// TwinCAT 3 PLC project otel
// Title: TcOtlp
// Company: S&E Engineering
// ProjectVersion: 0.0.0.1
// ProgramVersion: 3.1.4026.27
// libraries:
//   Tc2_Standard, * (Beckhoff Automation GmbH)
//   Tc2_System, * (Beckhoff Automation GmbH)
//   Tc2_Utilities, * (Beckhoff Automation GmbH)
//   Tc3_IotBase, * (Beckhoff Automation GmbH)
//   Tc3_JsonXml, * (Beckhoff Automation GmbH)
// project tree:
//   OTEL/COMMON/ENUMS/ E_BytesEncoding.TcTLEO
//   OTEL/COMMON/FUNCTION_BLOCKS/ FB_InstrumentationScope.TcPOU, FB_Resource.TcPOU
//   OTEL/COMMON/STRUCTS/ ST_LinkedListNode.TcDUT
//   OTEL/EXPORTING/ENUMS/ E_FileExporterState.TcTLEO, E_HttpExporterState.TcTLEO
//   OTEL/LOGGING/EXPORTING/ENUMS/ E_LogRecordExporterFailureReason.TcTLEO, E_LogRecordExporterState.TcTLEO
//   OTEL/LOGGING/EXPORTING/FUNCTION_BLOCKS/ FB_LogRecordExporter_Base.TcPOU, FB_LogRecordExporter_Console.TcPOU, FB_LogRecordExporter_File.TcPOU, FB_LogRecordExporter_HTTP.TcPOU
//   OTEL/LOGGING/LOGGER/ENUMS/ E_LoggerFailureReason.TcTLEO
//   OTEL/LOGGING/LOGGER/FUNCTION_BLOCKS/ FB_Logger.TcPOU
//   OTEL/LOGGING/LOG_RECORD/ENUMS/ E_LogRecordCloneFailureReason.TcTLEO, E_LogRecordFlag.TcTLEO, E_LogRecordQueueFailureReason.TcTLEO, E_SeverityNumber.TcTLEO
//   OTEL/LOGGING/LOG_RECORD/FUNCTION_BLOCKS/ FB_LogRecord.TcPOU, FB_LogRecordQueue.TcPOU
//   OTEL/LOGGING/PROCESSORS/ENUMS/ E_LogRecordProcessorFailureReason.TcTLEO
//   OTEL/LOGGING/PROCESSORS/FUNCTION_BLOCKS/ FB_LogRecordProcessor_Base.TcPOU, FB_LogRecordProcessor_Batch.TcPOU, FB_LogRecordProcessor_Simple.TcPOU
//   OTEL/LOGGING/PROVIDER/ENUMS/ E_LoggerProviderFailureReason.TcTLEO
//   OTEL/LOGGING/PROVIDER/FUNCTION_BLOCKS/ FB_LoggerProvider.TcPOU
//   OTEL/LOGGING/SERIALIZATION/FUNCTION_BLOCKS/ FB_LogRecordProtoJsonSerializer.TcPOU
//   OTEL/ TcOtlp_GVL.TcGVL
//   OTEL/TRACING/EXPORTING/ENUMS/ E_SpanExporterFailureReason.TcTLEO
//   OTEL/TRACING/EXPORTING/FUNCTION_BLOCKS/ FB_SpanExporter_Base.TcPOU, FB_SpanExporter_File.TcPOU, FB_SpanExporter_Console.TcPOU, FB_SpanExporter_HTTP.TcPOU
//   OTEL/TRACING/SPAN/ENUMS/ E_SpanCloneFailureReason.TcTLEO, E_SpanFlags.TcTLEO, E_ContextFactoryFailureReason.TcTLEO, E_SpanKind.TcTLEO, E_SpanQueueFailureReason.TcTLEO, E_StatusCode.TcTLEO
//   OTEL/TRACING/PROCESSORS/ENUMS/ E_SpanProcessorFailureReason.TcTLEO
//   OTEL/TRACING/PROCESSORS/FUNCTION_BLOCKS/ FB_SpanProcessor_Batch.TcPOU, FB_SpanProcessor_Base.TcPOU, FB_SpanProcessor_Simple.TcPOU
//   OTEL/EXPORTING/STRUCTS/ ST_HttpEndpoint.TcDUT
//   OTEL/EXPORTING/FUNCTIONS/ F_ParseHttpUrl.TcPOU
//   OTEL/TRACING/TRACESTATE/ENUMS/ E_TraceStateFailureReason.TcTLEO
//   OTEL/TRACING/TRACESTATE/FUNCTION_BLOCKS/ FB_TraceState.TcPOU, TraceStateFactory.TcPOU
//   OTEL/TRACING/PROPAGATION/ENUMS/ E_PropagationFailureReason.TcTLEO
//   OTEL/TRACING/PROPAGATION/ TraceContextPropagator.TcPOU
//   OTEL/TRACING/PROPAGATION/STRUCTS/ ST_TraceContextCarrier.TcDUT
//   OTEL/TRACING/SAMPLING/FUNCTION_BLOCKS/ FB_Sampler.TcPOU, FB_Sampler_AlwaysOn.TcPOU, FB_Sampler_ErrorsOnly.TcPOU
//   OTEL/TRACING/ID_GENERATION/ENUMS/ E_IdGenFailureReason.TcTLEO
//   OTEL/TRACING/ID_GENERATION/FUNCTION_BLOCKS/ FB_IdGenerator.TcPOU, FB_IdGenerator_Base.TcPOU
//   OTEL/TRACING/LINK/ENUM/ E_LinkFailureReason.TcTLEO
//   OTEL/TRACING/LINK/FUNCTION_BLOCKS/ FB_Link.TcPOU, FB_Links.TcPOU, LinkFactory.TcPOU
//   OTEL/TRACING/PROVIDER/ENUMS/ E_TracerProviderFailureReason.TcTLEO
//   OTEL/TRACING/PROVIDER/FUNCTION_BLOCKS/ FB_TracerProvider.TcPOU
//   OTEL/TRACING/SERIALIZATION/FUNCTION_BLOCKS/ FB_SpanProtoJsonSerializer.TcPOU
//   OTEL/TRACING/SPAN/ ContextFactory.TcPOU
//   OTEL/TRACING/SPAN/FUNCTION_BLOCKS/ FB_Span.TcPOU, FB_SpanContext.TcPOU, FB_SpanQueue.TcPOU, FB_Status.TcPOU
//   OTEL/TRACING/TRACER/ENUMS/ E_TracerFailureReason.TcTLEO
//   OTEL/TRACING/TRACER/ FB_Tracer.TcPOU
//   OTEL/VALUES/ENUMS/ E_AttributesFailureReason.TcTLEO, E_ValueFactoryFailureReason.TcTLEO, E_ValueType.TcTLEO
//   OTEL/VALUES/FUNCTION_BLOCKS/ FB_AnyValue.TcPOU, FB_Attributes.TcPOU, FB_KeyValue.TcPOU, FB_Number.TcPOU, FB_SpanId.TcPOU, FB_String.TcPOU, FB_TraceId.TcPOU
//   OTEL/VALUES/INTERFACES/ I_OtlpValue.TcIO
//   OTEL/VALUES/ ValueFactory.TcPOU
//   OTEL/SERIALIZATION/FUNCTION_BLOCKS/ FB_BaseProtoJsonSerializer.TcPOU
//   OTEL/SERIALIZATION/ENUMS/ E_ProtoJsonSerializerFailureReason.TcTLEO
//   Project Information/ F_GetCompany.TcPOU, F_GetTitle.TcPOU, F_GetVersion.TcPOU
//   Version/ Global_Version.TcGVL
// (motion and I/O tree: see PLC project test)
// real-time tasks:
//   TASK PlcTask: cycle T#10ms, priority 20, ADS port 350

// ---- OTEL/COMMON/ENUMS/E_BytesEncoding.TcTLEO
{attribute 'qualified_only'}
{attribute 'strict'}
{attribute 'to_string'}
TYPE E_BytesEncoding :
(
	hex := 0,
	base64
);
END_TYPE

// ---- OTEL/COMMON/STRUCTS/ST_LinkedListNode.TcDUT
{attribute 'enable_dynamic_creation'}
TYPE ST_LinkedListNode :
STRUCT
	val: PVOID;
	nxt: POINTER TO ST_LinkedListNode;
END_STRUCT
END_TYPE

// ---- OTEL/EXPORTING/ENUMS/E_FileExporterState.TcTLEO
{attribute 'qualified_only'}
{attribute 'strict'}
{attribute 'to_string'}
TYPE E_FileExporterState :
(
	error := -10,
	idle := 0,
	serializing := 10,
	creating := 15,
	opening := 20,
	buffering := 25,
	writing := 30,
	closing := 40,
	rotating := 50,
	done := 99
);
END_TYPE
//  error = '-10'

// ---- OTEL/EXPORTING/ENUMS/E_HttpExporterState.TcTLEO
{attribute 'qualified_only'}
{attribute 'strict'}
{attribute 'to_string'}
TYPE E_HttpExporterState :
(
	error := -10,
	idle := 0,
	serializing := 10,
	sending := 20,
	waiting := 30,
	processing := 40,
	done := 99
);
END_TYPE
//  error = '-10'

// ---- OTEL/LOGGING/EXPORTING/ENUMS/E_LogRecordExporterFailureReason.TcTLEO
{attribute 'qualified_only'}
{attribute 'strict'}
{attribute 'to_string'}
TYPE E_LogRecordExporterFailureReason :
(
	NA := 0,  // No failure occurred.
	ACTIVE_EXPORT_IN_PROGRESS,  // The exporter cannot accept another batch while an export is active.
	QUEUE_TRANSFER_FAILURE,  // Records could not be transferred into the exporter queue.
	SERIALIZATION_FAILURE,  // The accepted records could not be serialized.
	BUFFER_ALLOCATION_FAILURE,  // The serialized payload buffer could not be allocated.
	FILE_OPEN_FAILURE,  // The destination file could not be opened.
	FILE_WRITE_FAILURE,  // The serialized payload could not be written.
	FILE_CLOSE_FAILURE,  // The destination file could not be closed.
	HTTP_URL_PARSE_FAILURE,  // The configured endpoint URL could not be parsed.
	HTTP_REQUEST_FAILURE,  // The HTTP request could not be sent or completed.
	HTTP_STATUS_FAILURE  // The server responded with a non-success HTTP status code.
) UDINT;
END_TYPE

// ---- OTEL/LOGGING/EXPORTING/ENUMS/E_LogRecordExporterState.TcTLEO
{attribute 'qualified_only'}
{attribute 'strict'}
{attribute 'to_string'}
TYPE E_LogRecordExporterState :
(
	SUCCESS := 0,
	BUSY,
	FAILURE
);
END_TYPE

// ---- OTEL/LOGGING/LOGGER/ENUMS/E_LoggerFailureReason.TcTLEO
{attribute 'qualified_only'}
{attribute 'strict'}
{attribute 'to_string'}
TYPE E_LoggerFailureReason :
(
	NA := 0,  // No failure occurred.
	LOG_RECORD_ALREADY_STARTED,  // A record is already being built by this logger.
	LOG_RECORD_NOT_STARTED,  // No active record is available to modify or emit.
	EVENT_NAME_INVALID,  // The event name could not be copied into an owned value.
	BODY_VALUE_POINTER_NULL,  // The supplied body value pointer is null.
	BODY_VALUE_INVALID,  // The supplied body value could not be cloned.
	BODY_VALUE_TYPE_UNSUPPORTED,  // The supplied body value type is not supported.
	ATTRIBUTE_VALUE_INVALID,  // An attribute could not be created from the supplied value.
	ATTRIBUTE_VALUE_TYPE_UNSUPPORTED,  // The supplied attribute value type is not supported.
	ATTRIBUTE_COUNT_LIMIT_REACHED,  // The record cannot own another attribute.
	SPAN_ID_BYTES_POINTER_NULL,  // The supplied Span ID byte pointer is null.
	SPAN_ID_BYTE_COUNT_TOO_SMALL,  // The supplied Span ID buffer is shorter than eight bytes.
	SPAN_ID_INVALID,  // The supplied Span ID could not be copied.
	TRACE_ID_BYTES_POINTER_NULL,  // The supplied Trace ID byte pointer is null.
	TRACE_ID_BYTE_COUNT_TOO_SMALL,  // The supplied Trace ID buffer is shorter than sixteen bytes.
	TRACE_ID_INVALID,  // The supplied Trace ID could not be copied.
	SNAPSHOT_COPY_FAILURE,  // The resource or instrumentation-scope snapshot could not be copied.
	MEMORY_ALLOCATION_FAILURE,  // Dynamic memory allocation failed.
	TRANSFER_TO_PROVIDER_FAILURE  // Could not transfer ownership of the record to the provider
) UDINT;
END_TYPE

// ---- OTEL/LOGGING/LOG_RECORD/ENUMS/E_LogRecordCloneFailureReason.TcTLEO
{attribute 'qualified_only'}
{attribute 'strict'}
{attribute 'to_string'}
TYPE E_LogRecordCloneFailureReason :
(
	NA := 0,  // No failure occurred.
	DESTINATION_ALREADY_ASSIGNED,  // The clone destination pointer is already assigned.
	EVENT_NAME_INVALID,  // The source event name could not be cloned.
	TRACE_ID_INVALID,  // The source Trace ID could not be cloned.
	SPAN_ID_INVALID,  // The source Span ID could not be cloned.
	BODY_VALUE_INVALID,  // The source body could not be cloned.
	BODY_VALUE_TYPE_UNSUPPORTED,  // The source body contains an unsupported value type.
	RESOURCE_COPY_FAILURE,  // The resource snapshot could not be copied.
	SCOPE_COPY_FAILURE,  // The instrumentation-scope snapshot could not be copied.
	ATTRIBUTE_COPY_FAILURE,  // The record attributes could not be copied.
	MEMORY_ALLOCATION_FAILURE  // Dynamic memory allocation failed.
) UDINT;
END_TYPE

// ---- OTEL/LOGGING/LOG_RECORD/ENUMS/E_LogRecordFlag.TcTLEO
{attribute 'qualified_only'}
{attribute 'strict'}
{attribute 'to_string'}
TYPE E_LogRecordFlag:
(
	// The zero value for the enum. Should not be used for comparisons.
	// Instead use bitwise "and" with the appropriate mask as shown above.
	LOG_RECORD_FLAGS_DO_NOT_USE := 0,
	// Bits 0-7 are used for trace flags.
	LOG_RECORD_FLAGS_TRACE_FLAGS_MASK := 255 //0x000000FF;
) UDINT;
END_TYPE
//  LOG_RECORD_FLAGS_TRACE_FLAGS_MASK = '255 '

// ---- OTEL/LOGGING/LOG_RECORD/ENUMS/E_LogRecordQueueFailureReason.TcTLEO
{attribute 'qualified_only'}
{attribute 'strict'}
{attribute 'to_string'}
TYPE E_LogRecordQueueFailureReason :
(
	NA := 0,  // No failure occurred.
	RECORD_POINTER_NULL,  // The supplied log-record pointer is null.
	DESTINATION_ALREADY_ASSIGNED,  // The pop destination pointer is already assigned.
	QUEUE_EMPTY,  // The queue contains no record to pop.
	MAX_SIZE_ENFORCEMENT_FAILURE := 5,  // The bounded eviction loop could not restore the configured maximum size.
	DESTINATION_NOT_EMPTY,  // The transfer destination already owns records.
	DESTINATION_CAPACITY_TOO_SMALL,  // The transfer destination cannot hold every source record.
	SELF_TRANSFER_NOT_ALLOWED,  // A queue cannot transfer ownership to itself.
	MEMORY_ALLOCATION_FAILURE  // Dynamic node allocation failed.
) UDINT;
END_TYPE

// ---- OTEL/LOGGING/LOG_RECORD/ENUMS/E_SeverityNumber.TcTLEO
{attribute 'qualified_only'}
{attribute 'strict'}
{attribute 'to_string'}
TYPE E_SeverityNumber :
(
	UNSPECIFIED := 0,
	TRACE,
	TRACE2,
	TRACE3,
	TRACE4,
	DEBUG,
	DEBUG2,
	DEBUG3,
	DEBUG4,
	INFO,
	INFO2,
	INFO3,
	INFO4,
	WARN,
	WARN2,
	WARN3,
	WARN4,
	ERROR,
	ERROR2,
	ERROR3,
	ERROR4,
	FATAL,
	FATAL2,
	FATAL3,
	FATAL4
);
END_TYPE

// ---- OTEL/LOGGING/PROCESSORS/ENUMS/E_LogRecordProcessorFailureReason.TcTLEO
{attribute 'qualified_only'}
{attribute 'strict'}
{attribute 'to_string'}
TYPE E_LogRecordProcessorFailureReason :
(
	NA := 0,  // No failure occurred.
	RECORD_CLONE_FAILURE,  // The emitted record could not be cloned for retention.
	QUEUE_PUSH_FAILURE,  // The retained record could not be transferred into the queue.
	EXPORT_FAILURE  // The exporter did not accept the prepared batch.
) UDINT;
END_TYPE

// ---- OTEL/LOGGING/PROVIDER/ENUMS/E_LoggerProviderFailureReason.TcTLEO
{attribute 'qualified_only'}
{attribute 'strict'}
{attribute 'to_string'}
TYPE E_LoggerProviderFailureReason :
(
	NA := 0,  // No failure occurred.
	RECORD_POINTER_NULL,  // The supplied log record pointer is null.
	QUEUE_POP_FAILURE,  // A record could not be popped from the provider's queue during cyclical processing.
	STAGE_PROCESSOR_FAILURE,  // A processor could not be added to the internal linked list for some reason.
	UNEXPECTED_NULL_PROCESSOR_POINTER,  // A processor pointer was invalid when being accessed internally to the provider.
	UNEXPECTED_NULL_LINKED_LIST_NODE  // A processor linked list poitner was invalid when being accessed internally to the provider.
) UDINT;
END_TYPE

// ---- OTEL/TRACING/EXPORTING/ENUMS/E_SpanExporterFailureReason.TcTLEO
(* Why a span exporter refused a batch or could not deliver it. *)
{attribute 'qualified_only'}
{attribute 'strict'}
{attribute 'to_string'}
TYPE E_SpanExporterFailureReason :
(
	NA := 0,  // No failure occurred.
	ACTIVE_EXPORT_IN_PROGRESS,  // The exporter cannot accept another batch while an export is active.
	QUEUE_TRANSFER_FAILURE,  // Spans could not be transferred into the exporter queue.
	SERIALIZATION_FAILURE,  // The accepted spans could not be serialized.
	BUFFER_ALLOCATION_FAILURE,  // The serialized payload buffer could not be allocated.
	FILE_OPEN_FAILURE,  // The destination file could not be opened.
	FILE_WRITE_FAILURE,  // The serialized payload could not be written.
	FILE_CLOSE_FAILURE,  // The destination file could not be closed.
	HTTP_URL_PARSE_FAILURE,  // The configured endpoint URL could not be parsed.
	HTTP_REQUEST_FAILURE,  // The HTTP request could not be sent or completed.
	HTTP_STATUS_FAILURE  // The server responded with a non-success HTTP status code.
) UDINT;
END_TYPE

// ---- OTEL/TRACING/SPAN/ENUMS/E_SpanCloneFailureReason.TcTLEO
(* Why FB_Span.cloneTo could not copy a span. *)
{attribute 'qualified_only'}
{attribute 'strict'}
{attribute 'to_string'}
TYPE E_SpanCloneFailureReason :
(
	NA := 0,  // No failure occurred.
	DESTINATION_ALREADY_ASSIGNED,  // The destination pointer was not 0.
	MEMORY_ALLOCATION_FAILURE,  // Dynamic memory allocation failed.
	VALUE_COPY_FAILURE,  // The name, an identifier, the trace state or the status message could not be copied.
	ATTRIBUTE_COPY_FAILURE,  // The span attributes could not be copied.
	LINK_COPY_FAILURE,  // A span link could not be copied.
	RESOURCE_COPY_FAILURE,  // The resource could not be copied.
	SCOPE_COPY_FAILURE  // The instrumentation scope could not be copied.
) UDINT;
END_TYPE

// ---- OTEL/TRACING/PROCESSORS/ENUMS/E_SpanProcessorFailureReason.TcTLEO
(* Why a span processor could not keep or export an ended span. *)
{attribute 'qualified_only'}
{attribute 'strict'}
{attribute 'to_string'}
TYPE E_SpanProcessorFailureReason :
(
	NA := 0,  // No failure occurred.
	SPAN_CLONE_FAILURE,  // The ended span could not be cloned for retention.
	QUEUE_PUSH_FAILURE,  // The clone could not be pushed onto the queue.
	EXPORT_FAILURE  // The exporter did not accept the prepared batch.
) UDINT;
END_TYPE

// ---- OTEL/EXPORTING/STRUCTS/ST_HttpEndpoint.TcDUT
(* An HTTP endpoint split out of a URL by F_ParseHttpUrl. *)
TYPE ST_HttpEndpoint :
STRUCT
	useTls: BOOL;  // TRUE for https
	host: T_MaxString;
	port: UINT;  // the explicit port, or 80 for http and 443 for https
	path: T_MaxString := '/';  // starts with '/'
END_STRUCT
END_TYPE

// ---- OTEL/TRACING/TRACESTATE/ENUMS/E_TraceStateFailureReason.TcTLEO
(* Why TraceStateFactory could not produce a trace state. *)
{attribute 'qualified_only'}
{attribute 'strict'}
{attribute 'to_string'}
TYPE E_TraceStateFailureReason :
(
	NA := 0,  // No failure.
	DESTINATION_ALREADY_ASSIGNED,  // The destination pointer already holds a trace state.
	SOURCE_POINTER_NULL,  // The source trace state is missing or has been freed.
	HEADER_POINTER_NULL,  // The header pointer is 0.
	HEADER_TOO_LONG,  // The header is longer than TraceStateFactory.MAX_HEADER_LENGTH.
	INVALID_KEY,  // An entry has a key that does not follow the W3C key grammar.
	INVALID_VALUE,  // An entry has no '=' or a value that does not follow the W3C value grammar.
	DUPLICATE_KEY,  // Two entries have the same key.
	TOO_MANY_ENTRIES,  // The header has more than TraceStateFactory.MAX_ENTRIES entries.
	MEMORY_ALLOCATION_FAILURE  // The trace state could not be allocated.
) UDINT;
END_TYPE

// ---- OTEL/TRACING/PROPAGATION/ENUMS/E_PropagationFailureReason.TcTLEO
(* Why TraceContextPropagator could not extract a span context from a carrier, or inject one into it. *)
{attribute 'qualified_only'}
{attribute 'strict'}
{attribute 'to_string'}
TYPE E_PropagationFailureReason :
(
	NA := 0,  // No failure.
	DESTINATION_ALREADY_ASSIGNED,  // The destination pointer already holds a span context.
	TRACEPARENT_EMPTY,  // No traceparent arrived, so there is no context to extract.
	TRACEPARENT_LENGTH_INVALID,  // The traceparent is shorter than 55 characters, or longer for version 00.
	VERSION_INVALID,  // The version is not two lowercase hex digits, or is the reserved ff.
	DELIMITER_INVALID,  // A field is not followed by '-', or a future version's flags are followed by something else.
	TRACE_ID_INVALID,  // The trace id is not 32 lowercase hex digits, or is all zero.
	SPAN_ID_INVALID,  // The parent span id is not 16 lowercase hex digits, or is all zero.
	TRACE_FLAGS_INVALID,  // The trace flags are not two lowercase hex digits.
	MEMORY_ALLOCATION_FAILURE,  // The span context, or a shortened trace state, could not be allocated.
	CONTEXT_POINTER_NULL,  // inject was given no span context.
	CONTEXT_INVALID  // The span context has an all-zero trace id or span id, so there is nothing to propagate.
) UDINT;
END_TYPE

// ---- OTEL/TRACING/PROPAGATION/STRUCTS/ST_TraceContextCarrier.TcDUT
(*
	The W3C Trace Context headers of one call, written by TraceContextPropagator.inject and read
	by extract. It is the contract between the propagator and a transport: a transport moves the
	whole block, so the receiver never sees a traceparent beside a stale tracestate, and it knows
	nothing about the headers' format. The traceparent fits version 00, and the tracestate fits
	the 512 characters W3C asks every vendor to propagate.
*)
TYPE ST_TraceContextCarrier :
STRUCT
	traceparent: STRING(55);
	tracestate: STRING(512);  // '' when the context has no trace state
END_STRUCT
END_TYPE

// ---- OTEL/TRACING/ID_GENERATION/ENUMS/E_IdGenFailureReason.TcTLEO
{attribute 'qualified_only'}
{attribute 'strict'}
{attribute 'to_string'}
TYPE E_IdGenFailureReason :
(
	NA := 0,  // No failure occurred.
	NO_IDENTIFIERS_AVAILABLE,  // The ring held too few bytes; the caller must retry on a later cycle.
	GUID_SERVICE_FAILED,  // The TwinCAT GUID service reported an error while the ring was being refilled.
	MEMORY_ALLOCATION_FAILURE,  // The ring could not be allocated.
	INVALID_CONFIGUATION  // parameters used to configure the generator were not valid
) UDINT;
END_TYPE

// ---- OTEL/TRACING/LINK/ENUM/E_LinkFailureReason.TcTLEO
(* Why a LinkFactory or FB_Links call failed. *)
{attribute 'qualified_only'}
{attribute 'strict'}
{attribute 'to_string'}
TYPE E_LinkFailureReason :
(
	NA := 0,  // No failure occurred.
	DESTINATION_ALREADY_ASSIGNED,  // The destination pointer was not 0.
	CONTEXT_POINTER_NULL,  // The span context pointer is null.
	CONTEXT_INVALID,  // The span context has an all zero trace id or span id.
	SPAN_POINTER_NULL,  // The span pointer is null.
	LINK_POINTER_NULL,  // The link pointer is null.
	LINK_COUNT_LIMIT_REACHED,  // The collection already holds maxCount links; the link was dropped and counted.
	LINKS_EMPTY,  // The collection holds no links.
	MEMORY_ALLOCATION_FAILURE,  // Dynamic memory allocation failed.
	ATTRIBUTE_COPY_FAILURE  // The link attributes could not be copied.
) UDINT;
END_TYPE

// ---- OTEL/TRACING/PROVIDER/ENUMS/E_TracerProviderFailureReason.TcTLEO
(* Why FB_TracerProvider.tick failed. *)
{attribute 'qualified_only'}
{attribute 'strict'}
{attribute 'to_string'}
TYPE E_TracerProviderFailureReason :
(
	NA := 0,  // No failure occurred.
	QUEUE_POP_FAILURE,  // An ended span could not be popped from the provider queue.
	STAGE_PROCESSOR_FAILURE,  // A processor could not be added to the staged list.
	UNEXPECTED_NULL_PROCESSOR_POINTER,  // A staged processor pointer was null.
	UNEXPECTED_NULL_LINKED_LIST_NODE,  // The staged list was shorter than stagedProcessorCount.
	ID_GENERATOR_TICK_FAILURE  // The id generator could not advance.
) UDINT;
END_TYPE

// ---- OTEL/TRACING/SPAN/ENUMS/E_SpanFlags.TcTLEO
{attribute 'qualified_only'}
{attribute 'strict'}
{attribute 'to_string'}
TYPE E_SpanFlags :
(
	// The zero value for the enum. Should not be used for comparisons.
	// Instead use bitwise "and" with the appropriate mask as shown above.
	SPAN_FLAGS_DO_NOT_USE := 16#0,

	// Bits 0-7 are used for trace flags.
	SPAN_FLAGS_TRACE_FLAGS_MASK := 16#000000FF,

	// Bits 8 and 9 are used to indicate that the parent span or link span is remote.
	// Bit 8 (`HAS_IS_REMOTE`) indicates whether the value is known.
	// Bit 9 (`IS_REMOTE`) indicates whether the span or link is remote.
	SPAN_FLAGS_CONTEXT_HAS_IS_REMOTE_MASK := 16#00000100,
	SPAN_FLAGS_CONTEXT_IS_REMOTE_MASK := 16#00000200

  // Bits 10-31 are reserved for future use.
) UDINT;
END_TYPE
//  SPAN_FLAGS_DO_NOT_USE = '16#0'
//  SPAN_FLAGS_TRACE_FLAGS_MASK = '16#000000FF'
//  SPAN_FLAGS_CONTEXT_HAS_IS_REMOTE_MASK = '16#00000100'
//  SPAN_FLAGS_CONTEXT_IS_REMOTE_MASK = '16#00000200  '

// ---- OTEL/TRACING/SPAN/ENUMS/E_ContextFactoryFailureReason.TcTLEO
{attribute 'qualified_only'}
{attribute 'strict'}
{attribute 'to_string'}
TYPE E_ContextFactoryFailureReason :
(
	NA := 0,  // No failure occurred.
	DESTINATION_ALREADY_ASSIGNED,  // The destination pointer was already assigned when the operation began.
	TRACE_ID_POINTER_NULL,  // The trace ID pointer is null.
	SPAN_ID_POINTER_NULL,  // The span ID pointer is null.
	MEMORY_ALLOCATION_FAILURE,  // Dynamic memory allocation failed.
	SPAN_POINTER_NULL  // fromSpan was given a null span pointer.
);
END_TYPE

// ---- OTEL/TRACING/SPAN/ENUMS/E_SpanKind.TcTLEO
{attribute 'qualified_only'}
{attribute 'strict'}
{attribute 'to_string'}
TYPE E_SpanKind :
(
	// Unspecified. Do NOT use as default.
	// Implementations MAY assume SpanKind to be INTERNAL when receiving UNSPECIFIED.
	SPAN_KIND_UNSPECIFIED := 0,
	
	// Indicates that the span represents an internal operation within an application,
	// as opposed to an operation happening at the boundaries. Default value.
	SPAN_KIND_INTERNAL := 1,
	
	// Indicates that the span covers server-side handling of an RPC or other
	// remote network request.
	SPAN_KIND_SERVER := 2,
	
	// Indicates that the span describes a request to some remote service.
	SPAN_KIND_CLIENT := 3,
	
	// Indicates that the span describes a producer sending a message to a broker.
	// Unlike CLIENT and SERVER, there is often no direct critical path latency relationship
	// between producer and consumer spans. A PRODUCER span ends when the message was accepted
	// by the broker while the logical processing of the message might span a much longer time.
	SPAN_KIND_PRODUCER := 4,
	
	// Indicates that the span describes consumer receiving a message from a broker.
	// Like the PRODUCER kind, there is often no direct critical path latency relationship
	// between producer and consumer spans.
	SPAN_KIND_CONSUMER := 5
) UDINT;
END_TYPE

// ---- OTEL/TRACING/SPAN/ENUMS/E_SpanQueueFailureReason.TcTLEO
{attribute 'qualified_only'}
{attribute 'strict'}
{attribute 'to_string'}
TYPE E_SpanQueueFailureReason :
(
	NA := 0,  // No failure occurred.
	SPAN_POINTER_NULL,  // The supplied span pointer is null.
	DESTINATION_ALREADY_ASSIGNED,  // The pop destination pointer is already assigned.
	QUEUE_EMPTY,  // The queue contains no span to pop.
	MAX_SIZE_ENFORCEMENT_FAILURE,  // The bounded eviction loop could not restore the configured maximum size.
	MEMORY_ALLOCATION_FAILURE,  // Dynamic node allocation failed.
	SELF_TRANSFER_NOT_ALLOWED,  // transferTo was asked to move spans into the same queue.
	DESTINATION_NOT_EMPTY  // transferTo needs an empty destination queue.
) UDINT;
END_TYPE

// ---- OTEL/TRACING/SPAN/ENUMS/E_StatusCode.TcTLEO
{attribute 'qualified_only'}
{attribute 'strict'}
{attribute 'to_string'}
TYPE E_StatusCode :
(
	// The default status.
	STATUS_CODE_UNSET := 0,
	// The Span has been validated by an Application developer or Operator to 
	// have completed successfully.
	STATUS_CODE_OK := 1,
	// The Span contains an error.
	STATUS_CODE_ERROR := 2
) UDINT;
END_TYPE

// ---- OTEL/TRACING/TRACER/ENUMS/E_TracerFailureReason.TcTLEO
{attribute 'qualified_only'}
{attribute 'strict'}
{attribute 'to_string'}
TYPE E_TracerFailureReason :
(
	NA := 0,  // No failure occurred.
	SPAN_ALREADY_STARTED,  // startSpan was called while a span was still being built.
	SPAN_NOT_STARTED,  // No span is being built to modify or hand over.
	SPAN_NAME_EMPTY,  // The span name is empty.
	SPAN_KIND_UNSPECIFIED,  // SPAN_KIND_UNSPECIFIED was given; OTLP says not to use it.
	PARENT_CONTEXT_POINTER_NULL,  // The parent context pointer is null.
	PARENT_CONTEXT_INVALID,  // The parent context has an all zero trace id or span id.
	ATTRIBUTE_VALUE_INVALID,  // An attribute could not be created from the supplied value.
	ATTRIBUTE_VALUE_TYPE_UNSUPPORTED,  // The supplied attribute value type is not supported.
	ATTRIBUTE_COUNT_LIMIT_REACHED,  // The span cannot own another attribute.
	DESTINATION_ALREADY_ASSIGNED,  // The destination pointer was already assigned when build began.
	IDENTIFIERS_UNAVAILABLE,  // The id generator had no identifiers ready; retry on a later cycle.
	ID_GENERATION_FAILURE,  // The id generator failed for another reason.
	SNAPSHOT_COPY_FAILURE,  // The resource or instrumentation-scope snapshot could not be copied.
	MEMORY_ALLOCATION_FAILURE,  // Dynamic memory allocation failed.
	SPAN_POINTER_NULL,  // A method for a running span, such as endSpan, was given a null span pointer.
	TRANSFER_TO_PROVIDER_FAILURE,  // The provider could not queue the ended span, so it was released.
	LINK_CONTEXT_POINTER_NULL,  // addLink was given a null span context pointer.
	LINK_CONTEXT_INVALID,  // The linked context has an all zero trace id or span id.
	LINK_COUNT_LIMIT_REACHED,  // The span cannot own another link.
	PARENT_SPAN_POINTER_NULL,  // setParentUsingSpan was given a null span pointer.
	PARENT_SPAN_INVALID,  // The parent span has not been built, so it has no trace id or span id.
	SPAN_STATUS_ALREADY_SET,  // The span already has a status, and the first one set wins.
	SPAN_INVALID,  // The span has not been built, so it has no trace id or span id.
	LINK_POINTER_NULL  // pushSpanLink was given a null link pointer.
) UDINT;
END_TYPE

// ---- OTEL/VALUES/ENUMS/E_AttributesFailureReason.TcTLEO
{attribute 'qualified_only'}
{attribute 'strict'}
{attribute 'to_string'}
TYPE E_AttributesFailureReason :
(
	NA := 0,  // No attribute failure occurred.
	KV_POINTER_NULL,  // The supplied key-value pair pointer is null.
	KV_KEY_POINTER_NULL,  // The key-value pair has no key.
	KV_VALUE_POINTER_NULL,  // The key-value pair has no value.
	KV_VALUE_INVALID,  // The key-value pair contains an invalid value.
	KV_VALUE_TYPE_UNSUPPORTED,  // The key-value pair contains an unsupported value type.
	ATTRIBUTE_COUNT_LIMIT_REACHED,  // Adding a new key would exceed the configured attribute count limit.
	MEMORY_ALLOCATION_FAILURE,  // Dynamic memory allocation failed.
	KEY_NOT_FOUND  // The source collection has no attribute with the requested key.
) UDINT;
END_TYPE

// ---- OTEL/VALUES/ENUMS/E_ValueFactoryFailureReason.TcTLEO
{attribute 'qualified_only'}
{attribute 'strict'}
{attribute 'to_string'}
TYPE E_ValueFactoryFailureReason :
(
	NA := 0,  // No failure occurred.
	DESTINATION_ALREADY_ASSIGNED,  // The destination pointer was already assigned when the operation began.
	SOURCE_POINTER_NULL,  // The source pointer is null.
	NUMBER_VALUE_POINTER_NULL,  // The numeric value pointer is null.
	NUMBER_VALUE_SIZE_INVALID,  // The numeric value size is zero or negative.
	KEY_POINTER_NULL,  // The key pointer is null.
	VALUE_POINTER_NULL,  // The value pointer is null.
	STRING_POINTER_NULL,  // The string pointer is null.
	SPAN_ID_BYTES_POINTER_NULL,  // The Span ID byte-array pointer is null.
	SPAN_ID_BYTE_COUNT_TOO_SMALL,  // The supplied byte count is too small for a Span ID.
	TRACE_ID_BYTES_POINTER_NULL,  // The Trace ID byte-array pointer is null.
	TRACE_ID_BYTE_COUNT_TOO_SMALL,  // The supplied byte count is too small for a Trace ID.
	UNSUPPORTED_VALUE_TYPE,  // The source value type is not supported by the factory operation.
	MEMORY_ALLOCATION_FAILURE  // Dynamic memory allocation failed.
);
END_TYPE

// ---- OTEL/VALUES/ENUMS/E_ValueType.TcTLEO
{attribute 'qualified_only'}
{attribute 'strict'}
{attribute 'to_string'}
TYPE E_ValueType :
(
	E_String := 0,
	E_TraceId,
	E_SpanId,
	E_AnyValue,
	E_KeyValue,
	E_Number
);
END_TYPE

// ---- OTEL/SERIALIZATION/ENUMS/E_ProtoJsonSerializerFailureReason.TcTLEO
{attribute 'qualified_only'}
{attribute 'strict'}
{attribute 'to_string'}
TYPE E_ProtoJsonSerializerFailureReason :
(
	NA := 0,  // No failure occurred.
	JSON_VALUE_INVALID,  // The destination JSON value is invalid.
	JSON_OPERATION_FAILURE,  // The JSON DOM parser could not create or append a value.
	KEY_POINTER_NULL,  // The supplied member-key pointer is null.
	VALUE_POINTER_NULL,  // The supplied OTLP value pointer is null.
	LOG_RECORD_POINTER_NULL,  // The supplied log-record pointer is null.
	NUMBER_VALUE_POINTER_NULL,  // The numeric value does not point to its concrete value.
	UNSUPPORTED_VALUE_TYPE,  // The OTLP value type is not supported.
	UNSUPPORTED_NUMBER_TYPE,  // The IEC numeric type is not supported.
	BYTES_POINTER_NULL,  // The byte-array pointer is null.
	BYTE_COUNT_ZERO,  // No bytes were supplied for encoding.
	STRING_POINTER_NULL,  // The destination or source string pointer is null.
	STRING_BUFFER_TOO_SMALL,  // The encoded value does not fit in the destination string.
	UNSUPPORTED_BYTES_ENCODING,  // The requested byte encoding is not supported.
	ATTRIBUTE_COLLECTION_INCONSISTENT,  // The attribute count and linked values disagree.
	LOG_RECORD_COLLECTION_INCONSISTENT,  // The queue count and linked records disagree.
	QUEUE_TRANSFER_FAILURE,  // Ownership could not be transferred to the serializer queue.
	QUEUE_POP_FAILURE,  // An owned record could not be removed from the serializer queue.
	QUEUE_ROTATE_FAILURE,  // The serializer queue could not preserve grouping order.
	LOOP_LIMIT_EXCEEDED,  // Serialization could not complete within GVL.MAX_LOOP_COUNT.
	SPAN_POINTER_NULL,  // The supplied span pointer is null.
	SPAN_COLLECTION_INCONSISTENT,  // The span queue count and linked spans disagree.
	MEMORY_ALLOCATION_FAILURE  // A working buffer could not be allocated.
) UDINT;
END_TYPE

// ---- OTEL/TcOtlp_GVL.TcGVL
{attribute 'qualified_only'}
VAR_GLOBAL CONSTANT
	// Program/logic safety limits
	DEFAULT_MAX_ATTRIBUTE_COUNT: 	UDINT := 20;  	// Maximum attributes for FB_Attributes
	DEFAULT_MAX_LINK_COUNT:			UDINT := 128;	// Maximum links a span keeps, the OpenTelemetry default
	MAX_LOOP_COUNT:					UDINT := 20000; // Maximum iterations a for/while loop can have
	MAX_LOG_RECORDS_PER_SCAN: 		UDINT := 100;  	// Maximum number of log records that can be emitted per scan.
	MAX_SPAN_RECORDS_PER_SCAN:		UDINT := 100;	// Maximum number of spans that can be emitted per scan.
END_VAR
VAR_GLOBAL
	_ID: UDINT := 1;
	defaultSampler: FB_Sampler;  // ParentBased(root=AlwaysOn); stateless, so providers share it
END_VAR

// ---- Version/Global_Version.TcGVL
{attribute 'TcGenerated'}
{attribute 'no-analysis'}
{attribute 'linkalways'}
// This function has been automatically generated from the project information.
VAR_GLOBAL CONSTANT
	{attribute 'const_non_replaced'}
	stLibVersion_TcOtlp : ST_LibVersion := (iMajor := 0, iMinor := 0, iBuild := 0, iRevision := 1, nFlags := 0, sVersion := '0.0.0.1');
END_VAR

// ---- OTEL/VALUES/INTERFACES/I_OtlpValue.TcIO
INTERFACE I_OtlpValue

PROPERTY eType : E_ValueType
GET
END_GET
END_PROPERTY

// deallocates all data owned by the value without deleting the object itself.
METHOD free
END_METHOD

END_INTERFACE

// ---- OTEL/VALUES/FUNCTION_BLOCKS/FB_Attributes.TcPOU
(*
	Owned collection of OTLP key-value attributes used across telemetry domains.
*)
{attribute 'enable_dynamic_creation'}
FUNCTION_BLOCK FB_Attributes
VAR
	_head: POINTER TO ST_LinkedListNode;
	_tail: POINTER TO ST_LinkedListNode;
	_cursor: POINTER TO ST_LinkedListNode;
END_VAR
VAR_OUTPUT
	count: UDINT;
	maxCount: UDINT;
	droppedCount: UDINT;
END_VAR

(* The enforced bound: maxCount, held to MAX_LOOP_COUNT so free always reaches the end. *)
METHOD _capacity : UDINT
_capacity := MIN(THIS^.maxCount, TcOtlp_GVL.MAX_LOOP_COUNT);
END_METHOD

(* The node holding the attribute named key, or 0 when there is none. Does not move the next cursor. *)
METHOD _findNode : POINTER TO ST_LinkedListNode
VAR_INPUT
	key: T_MaxString;
END_VAR
VAR
	_idx: UDINT;
	_node: POINTER TO ST_LinkedListNode;
	_pKv: POINTER TO FB_KeyValue;
END_VAR
_findNode := 0;

_node := THIS^._head;
FOR _idx := 0 TO TcOtlp_GVL.MAX_LOOP_COUNT DO
	IF _node = 0 THEN
		RETURN;
	END_IF
	_pKv := _node^.val;
	IF _pKv <> 0 AND_THEN _pKv^.pKey <> 0 AND_THEN _pKv^.pKey^ = key THEN
		_findNode := _node;
		RETURN;
	END_IF
	_node := _node^.nxt;
END_FOR
END_METHOD

METHOD _mapValueFactoryFailure : E_AttributesFailureReason
VAR_INPUT
	failureReason: E_ValueFactoryFailureReason;
END_VAR
CASE failureReason OF
	E_ValueFactoryFailureReason.SOURCE_POINTER_NULL:
		_mapValueFactoryFailure := E_AttributesFailureReason.KV_VALUE_POINTER_NULL;
	E_ValueFactoryFailureReason.KEY_POINTER_NULL:
		_mapValueFactoryFailure := E_AttributesFailureReason.KV_KEY_POINTER_NULL;
	E_ValueFactoryFailureReason.VALUE_POINTER_NULL:
		_mapValueFactoryFailure := E_AttributesFailureReason.KV_VALUE_POINTER_NULL;
	E_ValueFactoryFailureReason.UNSUPPORTED_VALUE_TYPE:
		_mapValueFactoryFailure := E_AttributesFailureReason.KV_VALUE_TYPE_UNSUPPORTED;
	E_ValueFactoryFailureReason.MEMORY_ALLOCATION_FAILURE:
		_mapValueFactoryFailure := E_AttributesFailureReason.MEMORY_ALLOCATION_FAILURE;
	ELSE
		_mapValueFactoryFailure := E_AttributesFailureReason.KV_VALUE_INVALID;
END_CASE
END_METHOD

(*
	Adds a copy of src's attribute named key, stored under destKey, or under key when destKey is
	empty. An attribute already held under that name is replaced, as with setAttribute. src is
	left unchanged and may be this collection, so an attribute can be copied to a new name in place.
*)
METHOD copyAttribute : BOOL
VAR_IN_OUT
	src: FB_Attributes;
END_VAR
VAR_INPUT
	key: T_MaxString;
	destKey: T_MaxString := '';
END_VAR
VAR_OUTPUT
	failureReason: E_AttributesFailureReason;
END_VAR
VAR
	_pSrc: POINTER TO FB_KeyValue;
	_pDest: POINTER TO FB_KeyValue;
	_factoryFailureReason: E_ValueFactoryFailureReason;
END_VAR
copyAttribute := FALSE;
failureReason := E_AttributesFailureReason.NA;

_pSrc := src.getAttribute(key);
IF _pSrc = 0 THEN
	failureReason := E_AttributesFailureReason.KEY_NOT_FOUND;
	RETURN;
END_IF

IF destKey = '' THEN
	destKey := key;
END_IF

IF NOT ValueFactory.createKeyValue(
	pDest:=_pDest,
	pKey:=ADR(destKey),
	pVal:=_pSrc^.pVal,
	failureReason=>_factoryFailureReason
) THEN
	failureReason := THIS^._mapValueFactoryFailure(_factoryFailureReason);
	RETURN;
END_IF

copyAttribute := THIS^.setAttribute(pValue:=_pDest, failureReason=>failureReason);
// setAttribute only takes ownership on success; release a rejected value
IF _pDest <> 0 THEN
	_pDest^.delete(pSelf:=_pDest);
END_IF
END_METHOD

(*
	Adds a copy of every attribute in src, and carries src's droppedCount over, so the copy
	reports the same loss as the original.
*)
METHOD copyFrom : BOOL
VAR_IN_OUT
	src: FB_Attributes;
END_VAR
VAR_OUTPUT
	failureReason: E_AttributesFailureReason;
END_VAR
VAR
	_idx: UDINT;
	_pSrc: POINTER TO FB_KeyValue;
	_pDest: POINTER TO FB_KeyValue;
	_factoryFailureReason: E_ValueFactoryFailureReason;
END_VAR
copyFrom := FALSE;
failureReason := E_AttributesFailureReason.NA;

THIS^.droppedCount := THIS^.droppedCount + src.droppedCount;
src.reset();
FOR _idx := 0 TO TcOtlp_GVL.MAX_LOOP_COUNT DO
	_pSrc := src.next();
	IF _pSrc = 0 THEN
		copyFrom := failureReason = E_AttributesFailureReason.NA;
		RETURN;
	END_IF
	IF NOT ValueFactory.cloneKeyValue(pDest:=_pDest, pSrc:=_pSrc, failureReason=>_factoryFailureReason) THEN
		failureReason := THIS^._mapValueFactoryFailure(_factoryFailureReason);
		RETURN;
	END_IF
	IF NOT THIS^.setAttribute(pValue:=_pDest, failureReason=>failureReason) THEN
		IF _pDest <> 0 THEN
			_pDest^.delete(pSelf:=_pDest);
		END_IF
		RETURN;
	END_IF
END_FOR

copyFrom := failureReason = E_AttributesFailureReason.NA;
END_METHOD

METHOD FB_Exit : BOOL
VAR_INPUT
	bInCopyCode: BOOL;
END_VAR
IF NOT bInCopyCode THEN
	THIS^.free();
END_IF
END_METHOD

//FB_Init is always available implicitly and it is used primarily for initialization.
//The return value is not evaluated. For a specific influence, you can also declare the
//methods explicitly and provide additional code there with the standard initialization
//code. You can evaluate the return value.
METHOD FB_Init: BOOL
VAR_INPUT
    bInitRetains: BOOL; // TRUE: the retain variables are initialized (reset warm / reset cold)
    bInCopyCode: BOOL;  // TRUE: the instance will be copied to the copy code afterward (online change) 
	maxCount: UDINT := 20;  
END_VAR
THIS^.maxCount := maxCount;
END_METHOD

(*
	Releases every owned attribute. setAttribute holds count to MAX_LOOP_COUNT, so the loop
	always reaches the end, even if maxCount is lowered after attributes were added. If it ever
	stops early, the unreleased nodes stay in the collection and free returns FALSE, so a later
	call can finish the job.
*)
METHOD free : BOOL
VAR
	_idx: UDINT;
	_node: POINTER TO ST_LinkedListNode;
	_kv: POINTER TO FB_KeyValue;
END_VAR
FOR _idx := 0 TO TcOtlp_GVL.MAX_LOOP_COUNT DO
	IF THIS^._head = 0 THEN
		EXIT;
	END_IF

	_node := THIS^._head;
	THIS^._head := _node^.nxt;
	IF _node^.val <> 0 THEN
		_kv := _node^.val;
		_node^.val := 0;
		_kv^.delete(pSelf:=_kv);
	END_IF
	__DELETE(_node);
	_node := 0;
	IF THIS^.count > 0 THEN
		THIS^.count := THIS^.count - 1;
	END_IF
END_FOR

IF THIS^._head = 0 THEN
	THIS^._tail := 0;
	THIS^.count := 0;
END_IF
THIS^._cursor := THIS^._head;
free := THIS^._head = 0;
END_METHOD

(*
	Returns the attribute named key, or 0 when there is none. The collection keeps ownership: the
	pointer is borrowed and stays valid only until that attribute is replaced or the collection is
	freed. Does not move the next cursor.
*)
METHOD getAttribute : POINTER TO FB_KeyValue
VAR_INPUT
	key: T_MaxString;
END_VAR
VAR
	_node: POINTER TO ST_LinkedListNode;
END_VAR
getAttribute := 0;

_node := THIS^._findNode(key);
IF _node <> 0 THEN
	getAttribute := _node^.val;
END_IF
END_METHOD

METHOD next : POINTER TO FB_KeyValue
next := 0;

IF THIS^._cursor <> 0 THEN
	next := THIS^._cursor^.val;
	THIS^._cursor := THIS^._cursor^.nxt;
END_IF
END_METHOD

METHOD reset
THIS^._cursor := THIS^._head;
END_METHOD

METHOD setAttribute : BOOL
VAR_IN_OUT
	pValue: POINTER TO FB_KeyValue;
END_VAR
VAR_OUTPUT
	failureReason: E_AttributesFailureReason;
END_VAR
VAR
	_node: POINTER TO ST_LinkedListNode;
	_pVal: POINTER TO FB_KeyValue;
END_VAR
setAttribute := FALSE;
failureReason := E_AttributesFailureReason.NA;

IF pValue = 0 THEN
	failureReason := E_AttributesFailureReason.KV_POINTER_NULL;
	RETURN;
END_IF

IF pValue^.pKey = 0 THEN
	failureReason := E_AttributesFailureReason.KV_KEY_POINTER_NULL;
	RETURN;
END_IF

IF pValue^.pVal = 0 THEN
	failureReason := E_AttributesFailureReason.KV_VALUE_POINTER_NULL;
	RETURN;
END_IF

// replace the value if the key already exists
_node := THIS^._findNode(pValue^.pKey^);
IF _node <> 0 THEN
	_pVal := _node^.val;
	_pVal^.delete(pSelf:=_pVal);
	_node^.val := pValue;
	setAttribute := failureReason = E_AttributesFailureReason.NA;
	pValue := 0;
	RETURN;
END_IF

IF THIS^.count >= THIS^._capacity() THEN
	failureReason := E_AttributesFailureReason.ATTRIBUTE_COUNT_LIMIT_REACHED;
	THIS^.droppedCount := THIS^.droppedCount + 1;
	RETURN;
END_IF

// if it doesn't exist append the key-value pair
_node := __NEW(ST_LinkedListNode);
IF _node = 0 THEN
	failureReason := E_AttributesFailureReason.MEMORY_ALLOCATION_FAILURE;
	RETURN;
END_IF

_node^.val := pValue;
_node^.nxt := 0;

IF THIS^._tail = 0 THEN
	THIS^._head := _node;
	THIS^._cursor := _node;
ELSE
	THIS^._tail^.nxt := _node;
END_IF

THIS^._tail := _node;
THIS^.count := THIS^.count + 1;

// Ownership transfers only after the value has been linked successfully.
pValue := 0;
setAttribute := failureReason = E_AttributesFailureReason.NA;
END_METHOD

METHOD setNumberAttribute : BOOL
VAR_INPUT
	key: T_MaxString;
	value: ANY_NUM;
END_VAR
VAR_OUTPUT
	failureReason: E_AttributesFailureReason;
END_VAR
VAR
	_pKv: POINTER TO FB_KeyValue;
	_pNum: POINTER TO FB_Number;
	_factoryFailureReason: E_ValueFactoryFailureReason;
END_VAR
setNumberAttribute := FALSE;
failureReason := E_AttributesFailureReason.NA;

IF NOT ValueFactory.createNumber_AnyType(
	pDest:=_pNum,
	value:=value,
	failureReason=>_factoryFailureReason
) THEN
	failureReason := THIS^._mapValueFactoryFailure(_factoryFailureReason);
	RETURN;
END_IF

IF NOT ValueFactory.createKeyValue(
	pDest:=_pKv,
	pKey:=ADR(key),
	pVal:=_pNum,
	failureReason=>_factoryFailureReason
) THEN
	failureReason := THIS^._mapValueFactoryFailure(_factoryFailureReason);
	_pNum^.delete(pSelf:=_pNum);
	RETURN;
END_IF
_pNum^.delete(pSelf:=_pNum);  // clean up the _pNum as its cloned in createKeyValue

setNumberAttribute := THIS^.setAttribute(pValue:=_pKv, failureReason=>failureReason);
// setAttribute only takes ownership on success; release a rejected value
IF _pKv <> 0 THEN
	_pKv^.delete(pSelf:=_pKv);
END_IF
END_METHOD

METHOD setNumberAttribute_AnyType : BOOL
VAR_INPUT
	key: T_MaxString;
	value: AnyType;
END_VAR
VAR_OUTPUT
	failureReason: E_AttributesFailureReason;
END_VAR
VAR
	_pKv: POINTER TO FB_KeyValue;
	_pNum: POINTER TO FB_Number;
	_factoryFailureReason: E_ValueFactoryFailureReason;
END_VAR
setNumberAttribute_AnyType := FALSE;
failureReason := E_AttributesFailureReason.NA;

IF NOT ValueFactory.createNumber_AnyType(
	pDest:=_pNum,
	value:=value,
	failureReason=>_factoryFailureReason
) THEN
	failureReason := THIS^._mapValueFactoryFailure(_factoryFailureReason);
	RETURN;
END_IF

IF NOT ValueFactory.createKeyValue(
	pDest:=_pKv,
	pKey:=ADR(key),
	pVal:=_pNum,
	failureReason=>_factoryFailureReason
) THEN
	failureReason := THIS^._mapValueFactoryFailure(_factoryFailureReason);
	_pNum^.delete(pSelf:=_pNum);
	RETURN;
END_IF
_pNum^.delete(pSelf:=_pNum);  // clean up the _pNum as its cloned in createKeyValue

setNumberAttribute_AnyType := THIS^.setAttribute(pValue:=_pKv, failureReason=>failureReason);
// setAttribute only takes ownership on success; release a rejected value
IF _pKv <> 0 THEN
	_pKv^.delete(pSelf:=_pKv);
END_IF
END_METHOD

METHOD setStringAttribute : BOOL
VAR_INPUT
	key: T_MaxString;
	value: T_MaxString;
END_VAR
VAR_OUTPUT
	failureReason: E_AttributesFailureReason;
END_VAR
VAR
	_pKv: POINTER TO FB_KeyValue;
	_pStr: POINTER TO FB_String;
	_factoryFailureReason: E_ValueFactoryFailureReason;
END_VAR
setStringAttribute := FALSE;
failureReason := E_AttributesFailureReason.NA;

IF NOT ValueFactory.createString(
	pDest:=_pStr,
	pString:=ADR(value),
	failureReason=>_factoryFailureReason
) THEN
	failureReason := THIS^._mapValueFactoryFailure(_factoryFailureReason);
	RETURN;
END_IF

IF NOT ValueFactory.createKeyValue(
	pDest:=_pKv,
	pKey:=ADR(key),
	pVal:=_pStr,
	failureReason=>_factoryFailureReason
) THEN
	failureReason := THIS^._mapValueFactoryFailure(_factoryFailureReason);
	_pStr^.delete(pSelf:=_pStr);
	RETURN;
END_IF
_pStr^.delete(pSelf:=_pStr);  // clean up the _pStr as its cloned in createKeyValue

setStringAttribute := THIS^.setAttribute(pValue:=_pKv, failureReason=>failureReason);
// setAttribute only takes ownership on success; release a rejected value
IF _pKv <> 0 THEN
	_pKv^.delete(pSelf:=_pKv);
END_IF
END_METHOD

END_FUNCTION_BLOCK

// ---- OTEL/VALUES/FUNCTION_BLOCKS/FB_KeyValue.TcPOU
{attribute 'enable_dynamic_creation'}
FUNCTION_BLOCK FB_KeyValue IMPLEMENTS I_OtlpValue
VAR_OUTPUT
	pKey: POINTER TO STRING;
	pVal: POINTER TO FB_AnyValue;
END_VAR

(*
	Releases this value and clears the caller's pointer to it: call it as p^.delete(pSelf:=p).
	pSelf is cleared before the value is freed, so the caller never keeps a dangling pointer.
	A pointer to any other object is refused and left untouched, and nothing is released.
*)
METHOD delete : BOOL
VAR_IN_OUT
	pSelf: POINTER TO FB_KeyValue;
END_VAR
VAR
	_pThis: POINTER TO FB_KeyValue;
END_VAR
_pThis := THIS;
IF pSelf <> _pThis THEN
	RETURN;
END_IF

pSelf := 0;
__DELETE(_pThis);
delete := TRUE;
END_METHOD

PROPERTY eType : E_ValueType
GET
eType := E_ValueType.E_KeyValue;
END_GET
END_PROPERTY

//FB_Exit must be implemented explicitly. If there is an implementation, then the
//method is called before the controller removes the code of the function block instance
//(implicit call). The return value is not evaluated.
METHOD FB_Exit: BOOL
VAR_INPUT
    bInCopyCode: BOOL;  // TRUE: the exit method is called in order to leave the instance which will be copied afterwards (online change).  
END_VAR
THIS^.free();
END_METHOD

//FB_Init is always available implicitly and it is used primarily for initialization.
//The return value is not evaluated. For a specific influence, you can also declare the
//methods explicitly and provide additional code there with the standard initialization
//code. You can evaluate the return value.
METHOD FB_Init: BOOL
VAR_INPUT
    bInitRetains: BOOL; // TRUE: the retain variables are initialized (reset warm / reset cold)
    bInCopyCode: BOOL;  // TRUE: the instance will be copied to the copy code afterward (online change)
	pKey: POINTER TO STRING;
	pVal: POINTER TO FB_AnyValue;
END_VAR
(* Validation and allocation are handled by ValueFactory.createKeyValue. The
factory transfers ownership of both pointers only after every step succeeds. *)
THIS^.pKey := pKey;
THIS^.pVal := pVal;
END_METHOD

(* deallocates all data owned by the value without deleting the object itself.*)
METHOD free
IF THIS^.pKey <> 0 THEN
	__DELETE(THIS^.pKey);
	THIS^.pKey := 0;
END_IF
IF THIS^.pVal <> 0 THEN
	THIS^.pVal^.delete(pSelf:=THIS^.pVal);
END_IF
END_METHOD

END_FUNCTION_BLOCK

// ---- OTEL/VALUES/FUNCTION_BLOCKS/FB_AnyValue.TcPOU
FUNCTION_BLOCK ABSTRACT FB_AnyValue IMPLEMENTS I_OtlpValue

(*
	Releases this value and clears the caller's pointer to it: call it as p^.delete(pSelf:=p).
	pSelf is cleared before the value is freed, so the caller never keeps a dangling pointer.
	A pointer to any other object is refused and left untouched, and nothing is released.
*)
METHOD ABSTRACT delete : BOOL
VAR_IN_OUT
	pSelf: POINTER TO FB_AnyValue;
END_VAR
END_METHOD

PROPERTY ABSTRACT eType : E_ValueType
GET
END_GET
END_PROPERTY

(* deallocates all data owned by the value without deleting the object itself.*)
METHOD ABSTRACT free
END_METHOD

END_FUNCTION_BLOCK

// ---- OTEL/VALUES/ValueFactory.TcPOU
PROGRAM ValueFactory
VAR CONSTANT
	nSpanIdBytes: USINT := 8;
	nTraceIdBytes: USINT := 16;
END_VAR

METHOD cloneAnyValue : BOOL
VAR_IN_OUT
	pDest: POINTER TO FB_AnyValue;
END_VAR
VAR_INPUT
	pSrc: POINTER TO FB_AnyValue;
END_VAR
VAR_OUTPUT
	failureReason: E_ValueFactoryFailureReason;
END_VAR
VAR
	_type: E_ValueType;
END_VAR
cloneAnyValue := FALSE;
failureReason := E_ValueFactoryFailureReason.NA;

IF pDest <> 0 THEN
	failureReason := E_ValueFactoryFailureReason.DESTINATION_ALREADY_ASSIGNED;
	RETURN;
END_IF

IF pSrc = 0 THEN
	failureReason := E_ValueFactoryFailureReason.SOURCE_POINTER_NULL;
	RETURN;
END_IF

_type := pSrc^.eType;
CASE _type OF
	E_ValueType.E_String:
		cloneAnyValue := ValueFactory.cloneString(pDest:=pDest, pSrc:=pSrc, failureReason=>failureReason);
	E_ValueType.E_Number:
		cloneAnyValue := ValueFactory.cloneNumber(pDest:=pDest, pSrc:=pSrc, failureReason=>failureReason);
	E_ValueType.E_KeyValue:
		cloneAnyValue := ValueFactory.cloneKeyValue(pDest:=pDest, pSrc:=pSrc, failureReason=>failureReason);
	ELSE
		failureReason := E_ValueFactoryFailureReason.UNSUPPORTED_VALUE_TYPE;
END_CASE
END_METHOD

METHOD cloneKeyValue : BOOL
VAR_IN_OUT
	pDest: POINTER TO FB_KeyValue;
END_VAR
VAR_INPUT
	pSrc: POINTER TO FB_KeyValue;
END_VAR
VAR_OUTPUT
	failureReason: E_ValueFactoryFailureReason;
END_VAR
cloneKeyValue := FALSE;
failureReason := E_ValueFactoryFailureReason.NA;

IF pDest <> 0 THEN
	failureReason := E_ValueFactoryFailureReason.DESTINATION_ALREADY_ASSIGNED;
	RETURN;
END_IF

IF pSrc = 0 THEN
	failureReason := E_ValueFactoryFailureReason.SOURCE_POINTER_NULL;
	RETURN;
END_IF

cloneKeyValue := ValueFactory.createKeyValue(
	pDest:=pDest,
	pKey:=pSrc^.pKey,
	pVal:=pSrc^.pVal,
	failureReason=>failureReason
);
END_METHOD

METHOD cloneNumber : BOOL
VAR_IN_OUT
	pDest: POINTER TO FB_Number;
END_VAR
VAR_INPUT
	pSrc: POINTER TO FB_Number;
END_VAR
VAR_OUTPUT
	failureReason: E_ValueFactoryFailureReason;
END_VAR
VAR
	_value: AnyType;
	_pNew: POINTER TO FB_Number;
END_VAR
cloneNumber := FALSE;
failureReason := E_ValueFactoryFailureReason.NA;

IF pDest <> 0 THEN
	failureReason := E_ValueFactoryFailureReason.DESTINATION_ALREADY_ASSIGNED;
	RETURN;
END_IF

IF pSrc = 0 THEN
	failureReason := E_ValueFactoryFailureReason.SOURCE_POINTER_NULL;
	RETURN;
END_IF

IF pSrc^.value.pValue = 0 THEN
	failureReason := E_ValueFactoryFailureReason.NUMBER_VALUE_POINTER_NULL;
	RETURN;
END_IF

IF pSrc^.value.diSize <= 0 THEN
	failureReason := E_ValueFactoryFailureReason.NUMBER_VALUE_SIZE_INVALID;
	RETURN;
END_IF

// because it's really verbose to extract the number back out of the number we manually clone numbers
_value := pSrc^.value;
_value.pValue := __NEW(BYTE, _value.diSize);
IF _value.pValue = 0 THEN
	failureReason := E_ValueFactoryFailureReason.MEMORY_ALLOCATION_FAILURE;
	RETURN;
END_IF
MEMCPY(_value.pValue, pSrc^.value.pValue, TO_UDINT(_value.diSize));

_pNew := __NEW(FB_Number(
	value:=_value
));
IF _pNew = 0 THEN
	failureReason := E_ValueFactoryFailureReason.MEMORY_ALLOCATION_FAILURE;
	__DELETE(_value.pValue);
	_value.pValue := 0;
	RETURN;
END_IF
_value.pValue := 0;  // moved into FB_Number
pDest := _pNew;
cloneNumber := failureReason = E_ValueFactoryFailureReason.NA;
END_METHOD

METHOD cloneString : BOOL
VAR_IN_OUT
	pDest: POINTER TO FB_String;
END_VAR
VAR_INPUT
	pSrc: POINTER TO FB_String;
END_VAR
VAR_OUTPUT
	failureReason: E_ValueFactoryFailureReason;
END_VAR
cloneString := FALSE;
failureReason := E_ValueFactoryFailureReason.NA;

IF pDest <> 0 THEN
	failureReason := E_ValueFactoryFailureReason.DESTINATION_ALREADY_ASSIGNED;
	RETURN;
END_IF

IF pSrc = 0 THEN
	failureReason := E_ValueFactoryFailureReason.SOURCE_POINTER_NULL;
	RETURN;
END_IF

IF pSrc^.pString = 0 THEN
	failureReason := E_ValueFactoryFailureReason.STRING_POINTER_NULL;
	RETURN;
END_IF

cloneString := ValueFactory.createString(pDest:=pDest, pString:=pSrc^.pString, failureReason=>failureReason);
END_METHOD

METHOD createKeyValue : BOOL
VAR_IN_OUT
	pDest: POINTER TO FB_KeyValue;
END_VAR
VAR_INPUT
	pKey: POINTER TO STRING;
	pVal: POINTER TO FB_AnyValue;
END_VAR
VAR_OUTPUT
	failureReason: E_ValueFactoryFailureReason;
END_VAR
VAR
	_pNew: POINTER TO FB_KeyValue;
	_pKey: POINTER TO STRING;
	_pVal: POINTER TO FB_AnyValue;
	_len: UDINT;
END_VAR
createKeyValue := FALSE;
failureReason := E_ValueFactoryFailureReason.NA;

IF pKey = 0 THEN
	failureReason := E_ValueFactoryFailureReason.KEY_POINTER_NULL;
	RETURN;
END_IF

IF pVal = 0 THEN
	failureReason := E_ValueFactoryFailureReason.VALUE_POINTER_NULL;
	RETURN;
END_IF

IF pDest <> 0 THEN
	failureReason := E_ValueFactoryFailureReason.DESTINATION_ALREADY_ASSIGNED;
	RETURN;
END_IF

// clone all owned data before allocating the value itself
_len := LEN2(pKey) + 1;
_pKey := __NEW(BYTE, _len);
IF _pKey = 0 THEN
	failureReason := E_ValueFactoryFailureReason.MEMORY_ALLOCATION_FAILURE;
	RETURN;
END_IF
MEMCPY(_pKey, pKey, _len);

createKeyValue := ValueFactory.cloneAnyValue(pDest:=_pVal, pSrc:=pVal, failureReason=>failureReason);
IF NOT createKeyValue THEN
	__DELETE(_pKey);
	_pKey := 0;
	IF _pVal <> 0 THEN _pVal^.delete(pSelf:=_pVal); END_IF
	RETURN;
END_IF

_pNew := __NEW(FB_KeyValue(pKey:=_pKey, pVal:=_pVal));
IF _pNew = 0 THEN
	createKeyValue := FALSE;
	failureReason := E_ValueFactoryFailureReason.MEMORY_ALLOCATION_FAILURE;
	__DELETE(_pKey);
	_pKey := 0;
	_pVal^.delete(pSelf:=_pVal);
	RETURN;
END_IF
_pKey := 0;  // moved into FB_KeyValue
_pVal := 0;
pDest := _pNew;
createKeyValue := failureReason = E_ValueFactoryFailureReason.NA;
END_METHOD

METHOD createNumber : BOOL
VAR_IN_OUT
	pDest: POINTER TO FB_Number;
END_VAR
VAR_INPUT
	value: ANY_NUM;
END_VAR
VAR_OUTPUT
	failureReason: E_ValueFactoryFailureReason;
END_VAR
createNumber := FALSE;
failureReason := E_ValueFactoryFailureReason.NA;

createNumber := ValueFactory.createNumber_AnyType(
	pDest:=pDest,
	value:=value,
	failureReason=>failureReason
);
END_METHOD

(*
	This method is necessary because it makes it possible to easily create
	instance of an FB_Number from already instantiated instances of FB_Number
	i.e. cloning, when the original number is gone, but the AnyType value exists.
*)
METHOD createNumber_AnyType : BOOL
VAR_IN_OUT
	pDest: POINTER TO FB_Number;
END_VAR
VAR_INPUT
	value: AnyType;  // notice this is a struct and not the ANY_NUM keyword
END_VAR
VAR_OUTPUT
	failureReason: E_ValueFactoryFailureReason;
END_VAR
VAR
	_value: AnyType;
	_pNew: POINTER TO FB_Number;
END_VAR
createNumber_AnyType := FALSE;
failureReason := E_ValueFactoryFailureReason.NA;

IF pDest <> 0 THEN
	failureReason := E_ValueFactoryFailureReason.DESTINATION_ALREADY_ASSIGNED;
	RETURN;
END_IF

IF value.pValue = 0 THEN
	failureReason := E_ValueFactoryFailureReason.NUMBER_VALUE_POINTER_NULL;
	RETURN;
END_IF

IF value.diSize <= 0 THEN
	failureReason := E_ValueFactoryFailureReason.NUMBER_VALUE_SIZE_INVALID;
	RETURN;
END_IF

// Copy the concrete numeric value so the wrapper never retains caller-owned data.
_value.TypeClass := value.TypeClass;
_value.diSize := value.diSize;
_value.pValue := __NEW(BYTE, TO_UDINT(_value.diSize));
IF _value.pValue = 0 THEN
	failureReason := E_ValueFactoryFailureReason.MEMORY_ALLOCATION_FAILURE;
	RETURN;
END_IF
MEMCPY(_value.pValue, value.pValue, TO_UDINT(value.diSize));

_pNew := __NEW(FB_Number(value:=_value));
IF _pNew = 0 THEN
	failureReason := E_ValueFactoryFailureReason.MEMORY_ALLOCATION_FAILURE;
	__DELETE(_value.pValue);
	_value.pValue := 0;
	RETURN;
END_IF
_value.pValue := 0;  // moved into FB_Number
pDest := _pNew;
createNumber_AnyType := failureReason = E_ValueFactoryFailureReason.NA;
END_METHOD

METHOD createSpanId : BOOL
VAR_IN_OUT
	pDest: POINTER TO FB_SpanId;
END_VAR
VAR_INPUT
	pBytes: POINTER TO BYTE;
	nSize: UDINT;
END_VAR
VAR_OUTPUT
	failureReason: E_ValueFactoryFailureReason;
END_VAR
VAR
	_pNew: POINTER TO FB_SpanId;
END_VAR
createSpanId := FALSE;
failureReason := E_ValueFactoryFailureReason.NA;

IF pDest <> 0 THEN
	failureReason := E_ValueFactoryFailureReason.DESTINATION_ALREADY_ASSIGNED;
	RETURN;
END_IF

IF pBytes = 0 THEN
	failureReason := E_ValueFactoryFailureReason.SPAN_ID_BYTES_POINTER_NULL;
	RETURN;
END_IF

IF nSize < ValueFactory.nSpanIdBytes THEN
	failureReason := E_ValueFactoryFailureReason.SPAN_ID_BYTE_COUNT_TOO_SMALL;
	RETURN;
END_IF

_pNew := __NEW(FB_SpanId);
IF _pNew = 0 THEN
	failureReason := E_ValueFactoryFailureReason.MEMORY_ALLOCATION_FAILURE;
	RETURN;
END_IF

MEMCPY(ADR(_pNew^.bytes), pBytes, SIZEOF(_pNew^.bytes));
pDest := _pNew;
createSpanId := failureReason = E_ValueFactoryFailureReason.NA;
END_METHOD

METHOD createString : BOOL
VAR_IN_OUT
	pDest: POINTER TO FB_String;
END_VAR
VAR_INPUT
	pString: POINTER TO STRING;
END_VAR
VAR_OUTPUT
	failureReason: E_ValueFactoryFailureReason;
END_VAR
VAR
	_pString: POINTER TO STRING;
	_pNew: POINTER TO FB_String;
	_len: UDINT;
END_VAR
createString := FALSE;
failureReason := E_ValueFactoryFailureReason.NA;

IF pDest <> 0  THEN
	failureReason := E_ValueFactoryFailureReason.DESTINATION_ALREADY_ASSIGNED;
	RETURN;
END_IF

IF pString = 0 THEN
	failureReason := E_ValueFactoryFailureReason.STRING_POINTER_NULL;
	RETURN;
END_IF

// clone the string into a new pointer so as to not use mutable data
// an extra character is needed for the terminating character, which is a literal 0 just like "cstrings"
_len := LEN2(pString) + 1;
_pString := __NEW(BYTE, _len);
IF _pString = 0 THEN
	failureReason := E_ValueFactoryFailureReason.MEMORY_ALLOCATION_FAILURE;
	RETURN;
END_IF
MEMCPY(_pString, pString, _len);

_pNew := __NEW(FB_String(pString:=_pString));
IF _pNew = 0 THEN
	failureReason := E_ValueFactoryFailureReason.MEMORY_ALLOCATION_FAILURE;
	__DELETE(_pString);
	_pString := 0;
	RETURN;
END_IF
_pString := 0;  // moved into FB_String
pDest := _pNew;
createString := failureReason = E_ValueFactoryFailureReason.NA;
END_METHOD

METHOD createTraceId : BOOL
VAR_IN_OUT
	pDest: POINTER TO FB_TraceId;
END_VAR
VAR_INPUT
	pBytes: POINTER TO BYTE;
	nSize: UDINT;
END_VAR
VAR_OUTPUT
	failureReason: E_ValueFactoryFailureReason;
END_VAR
VAR
	_pNew: POINTER TO FB_TraceId;
END_VAR
createTraceId := FALSE;
failureReason := E_ValueFactoryFailureReason.NA;

IF pDest <> 0 THEN
	failureReason := E_ValueFactoryFailureReason.DESTINATION_ALREADY_ASSIGNED;
	RETURN;
END_IF

IF pBytes = 0 THEN
	failureReason := E_ValueFactoryFailureReason.TRACE_ID_BYTES_POINTER_NULL;
	RETURN;
END_IF

IF nSize < ValueFactory.nTraceIdBytes THEN
	failureReason := E_ValueFactoryFailureReason.TRACE_ID_BYTE_COUNT_TOO_SMALL;
	RETURN;
END_IF

_pNew := __NEW(FB_TraceId);
IF _pNew = 0 THEN
	failureReason := E_ValueFactoryFailureReason.MEMORY_ALLOCATION_FAILURE;
	RETURN;
END_IF
MEMCPY(ADR(_pNew^.bytes), pBytes, SIZEOF(_pNew^.bytes));
pDest := _pNew;
createTraceId := failureReason = E_ValueFactoryFailureReason.NA;
END_METHOD

END_PROGRAM

// ---- OTEL/VALUES/FUNCTION_BLOCKS/FB_Number.TcPOU
{attribute 'enable_dynamic_creation'}
FUNCTION_BLOCK FB_Number EXTENDS FB_AnyValue IMPLEMENTS I_OtlpValue
VAR_OUTPUT
	value: AnyType;
END_VAR

(*
	Releases this value and clears the caller's pointer to it: call it as p^.delete(pSelf:=p).
	pSelf is cleared before the value is freed, so the caller never keeps a dangling pointer.
	A pointer to any other object is refused and left untouched, and nothing is released.
*)
METHOD delete : BOOL
VAR_IN_OUT
	pSelf: POINTER TO FB_AnyValue;
END_VAR
VAR
	_pThis: POINTER TO FB_Number;
	_pSelfAsParam: POINTER TO FB_AnyValue;
END_VAR
_pThis := THIS;
_pSelfAsParam := _pThis;
IF pSelf <> _pSelfAsParam THEN
	RETURN;
END_IF

pSelf := 0;
__DELETE(_pThis);
delete := TRUE;
END_METHOD

PROPERTY eType : E_ValueType
GET
eType := E_ValueType.E_Number;
END_GET
END_PROPERTY

//FB_Exit must be implemented explicitly. If there is an implementation, then the
//method is called before the controller removes the code of the function block instance
//(implicit call). The return value is not evaluated.
METHOD FB_Exit: BOOL
VAR_INPUT
    bInCopyCode: BOOL;  // TRUE: the exit method is called in order to leave the instance which will be copied afterwards (online change).  
END_VAR
THIS^.free();
END_METHOD

//FB_Init is always available implicitly and it is used primarily for initialization.
//The return value is not evaluated. For a specific influence, you can also declare the
//methods explicitly and provide additional code there with the standard initialization
//code. You can evaluate the return value.
METHOD FB_Init: BOOL
VAR_INPUT
    bInitRetains: BOOL; // TRUE: the retain variables are initialized (reset warm / reset cold)
    bInCopyCode: BOOL;  // TRUE: the instance will be copied to the copy code afterward (online change)
	value: AnyType;
END_VAR
(* ValueFactory owns validation and allocation. FB_Number takes ownership of
the copied value and its type metadata only after every allocation succeeds. *)
THIS^.value := value;
END_METHOD

(* deallocates all data owned by the value without deleting the object itself.*)
METHOD free
IF THIS^.value.pValue <> 0 THEN
	__DELETE(THIS^.value.pValue);
END_IF
MEMSET(ADR(THIS^.value), 0, SIZEOF(THIS^.value));
END_METHOD

END_FUNCTION_BLOCK

// ---- OTEL/VALUES/FUNCTION_BLOCKS/FB_String.TcPOU
{attribute 'enable_dynamic_creation'}
FUNCTION_BLOCK FB_String EXTENDS FB_AnyValue IMPLEMENTS I_OtlpValue
VAR_OUTPUT
	pString: POINTER TO STRING;
END_VAR

(*
	Releases this value and clears the caller's pointer to it: call it as p^.delete(pSelf:=p).
	pSelf is cleared before the value is freed, so the caller never keeps a dangling pointer.
	A pointer to any other object is refused and left untouched, and nothing is released.
*)
METHOD delete : BOOL
VAR_IN_OUT
	pSelf: POINTER TO FB_AnyValue;
END_VAR
VAR
	_pThis: POINTER TO FB_String;
	_pSelfAsParam: POINTER TO FB_AnyValue;
END_VAR
_pThis := THIS;
_pSelfAsParam := _pThis;
IF pSelf <> _pSelfAsParam THEN
	RETURN;
END_IF

pSelf := 0;
__DELETE(_pThis);
delete := TRUE;
END_METHOD

PROPERTY eType : E_ValueType
GET
eType := E_ValueType.E_String;
END_GET
END_PROPERTY

//FB_Exit must be implemented explicitly. If there is an implementation, then the
//method is called before the controller removes the code of the function block instance
//(implicit call). The return value is not evaluated.
METHOD FB_Exit: BOOL
VAR_INPUT
    bInCopyCode: BOOL;  // TRUE: the exit method is called in order to leave the instance which will be copied afterwards (online change).  
END_VAR
THIS^.free();
END_METHOD

//FB_Init is always available implicitly and it is used primarily for initialization.
//The return value is not evaluated. For a specific influence, you can also declare the
//methods explicitly and provide additional code there with the standard initialization
//code. You can evaluate the return value.
METHOD FB_Init: BOOL
VAR_INPUT
    bInitRetains: BOOL; // TRUE: the retain variables are initialized (reset warm / reset cold)
    bInCopyCode: BOOL;  // TRUE: the instance will be copied to the copy code afterward (online change)
	pString: POINTER TO STRING;
END_VAR
(* 
Allocation and validation of the bytes is done at the
ValueFactory and not the value iteself, that way a new value 
never gets allocated if the initialization fails.
*)
THIS^.pString := pString;
END_METHOD

METHOD free
IF THIS^.pString <> 0 THEN
	__DELETE(THIS^.pString);
	THIS^.pString := 0;
END_IF
END_METHOD

END_FUNCTION_BLOCK

// ---- OTEL/VALUES/FUNCTION_BLOCKS/FB_SpanId.TcPOU
{attribute 'enable_dynamic_creation'}
FUNCTION_BLOCK FB_SpanId IMPLEMENTS I_OtlpValue
VAR_OUTPUT
	bytes: ARRAY [0..7] OF BYTE;
END_VAR

(*
	Releases this value and clears the caller's pointer to it: call it as p^.delete(pSelf:=p).
	pSelf is cleared before the value is freed, so the caller never keeps a dangling pointer.
	A pointer to any other object is refused and left untouched, and nothing is released.
*)
METHOD delete : BOOL
VAR_IN_OUT
	pSelf: POINTER TO FB_SpanId;
END_VAR
VAR
	_pThis: POINTER TO FB_SpanId;
END_VAR
_pThis := THIS;
IF pSelf <> _pThis THEN
	RETURN;
END_IF

pSelf := 0;
__DELETE(_pThis);
delete := TRUE;
END_METHOD

PROPERTY eType : E_ValueType
GET
eType := E_ValueType.E_SpanId;
END_GET
END_PROPERTY

//FB_Exit must be implemented explicitly. If there is an implementation, then the
//method is called before the controller removes the code of the function block instance
//(implicit call). The return value is not evaluated.
METHOD FB_Exit: BOOL
VAR_INPUT
    bInCopyCode: BOOL;  // TRUE: the exit method is called in order to leave the instance which will be copied afterwards (online change).  
END_VAR
THIS^.free();
END_METHOD

(* deallocates all data owned by the value without deleting the object itself.*)
METHOD free
MEMSET(ADR(THIS^.bytes), 0, SIZEOF(THIS^.bytes));
END_METHOD

END_FUNCTION_BLOCK

// ---- OTEL/VALUES/FUNCTION_BLOCKS/FB_TraceId.TcPOU
{attribute 'enable_dynamic_creation'}
FUNCTION_BLOCK FB_TraceId IMPLEMENTS I_OtlpValue
VAR_OUTPUT
	bytes: ARRAY [0..15] OF BYTE;
END_VAR

(*
	Releases this value and clears the caller's pointer to it: call it as p^.delete(pSelf:=p).
	pSelf is cleared before the value is freed, so the caller never keeps a dangling pointer.
	A pointer to any other object is refused and left untouched, and nothing is released.
*)
METHOD delete : BOOL
VAR_IN_OUT
	pSelf: POINTER TO FB_TraceId;
END_VAR
VAR
	_pThis: POINTER TO FB_TraceId;
END_VAR
_pThis := THIS;
IF pSelf <> _pThis THEN
	RETURN;
END_IF

pSelf := 0;
__DELETE(_pThis);
delete := TRUE;
END_METHOD

PROPERTY eType : E_ValueType
GET
eType := E_ValueType.E_TraceId;
END_GET
END_PROPERTY

//FB_Exit must be implemented explicitly. If there is an implementation, then the
//method is called before the controller removes the code of the function block instance
//(implicit call). The return value is not evaluated.
METHOD FB_Exit: BOOL
VAR_INPUT
    bInCopyCode: BOOL;  // TRUE: the exit method is called in order to leave the instance which will be copied afterwards (online change).  
END_VAR
THIS^.free();
END_METHOD

METHOD free
// just resets values to defaults
MEMSET(ADR(THIS^.bytes), 0, SIZEOF(THIS^.bytes));
END_METHOD

END_FUNCTION_BLOCK

// ---- OTEL/TRACING/SAMPLING/FUNCTION_BLOCKS/FB_Sampler.TcPOU
(*
	Decides which spans are sampled, through the sampled bit of the span's trace flags. The
	tracer calls onStart when it builds a span, and FB_TracerProvider calls onEnd when the span
	ends. A span is processed only if its sampled bit is still set after both.

	Used as is, this is the OpenTelemetry default ParentBased(root=AlwaysOn): a root span is
	sampled, and a child keeps its parent's decision, including a remote parent's. Extend it and
	override either method to change the policy:
	  onStart - the head decision. It can set or clear the bit, and the bit is carried into the
	            span's context, so children and injected carriers inherit it.
	  onEnd   - a later decision, made once the span's status is known. The provider calls it only
	            for spans that are still sampled, so it can drop a span but never keep one that
	            onStart dropped.
	Both methods borrow the span for the call and must not keep it.
*)
FUNCTION_BLOCK FB_Sampler

(* Samples a root span; a child keeps the sampled bit it copied from its parent. *)
METHOD onStart
VAR_INPUT
	span: REFERENCE TO FB_Span;
END_VAR
IF span.parentSpanId = 0 THEN
	span.setSampled(TRUE);
END_IF
END_METHOD

(* Keeps every span that is still sampled. *)
METHOD onEnd
VAR_INPUT
	span: REFERENCE TO FB_Span;
END_VAR
END_METHOD

END_FUNCTION_BLOCK

// ---- OTEL/TRACING/SPAN/FUNCTION_BLOCKS/FB_Span.TcPOU
(*
	One timed operation in a trace. Unlike a log record, a span has a lifecycle:
	  building - FB_Tracer owns it while the fluent chain fills it in,
	  running  - build hands it to the caller, who owns it while the work runs,
	  ended    - FB_Tracer.endSpan hands it to the provider for processing.
	The span owns every pointer member and releases them in free. A running span is read and
	changed only through FB_Tracer, such as getSpanContext, setSpanStatusOk and discardSpan,
	so callers never dereference it themselves. The methods left here belong to the tracing
	pipeline: the provider, samplers and processors.
*)
{attribute 'enable_dynamic_creation'}
FUNCTION_BLOCK FB_Span
VAR_INPUT
	// written by the tracer while the span is built
	name: POINTER TO FB_String;
	kind: E_SpanKind;
	startTimestamp: ULINT;
	endTimestamp: ULINT;
	traceId: POINTER TO FB_TraceId;
	spanId: POINTER TO FB_SpanId;
	traceState: POINTER TO FB_TraceState;

	// required if child span, must be omitted if root span
	parentSpanId: POINTER TO FB_SpanId;

	// describes the parent's remoteness, not this span's; see E_SpanFlags
	flags: UDINT;
	status: POINTER TO FB_Status;
END_VAR
VAR_OUTPUT
	attributes: FB_Attributes(maxCount := TcOtlp_GVL.DEFAULT_MAX_ATTRIBUTE_COUNT);
	links: FB_Links(maxCount := TcOtlp_GVL.DEFAULT_MAX_LINK_COUNT);
	resource: FB_Resource('');
	scope: FB_InstrumentationScope('', '', '');

	// span events have been deprecated, instead logs should be emitted with span context for correlation
	// events
	// droppedEventCount
END_VAR

(*
	Releases this span and clears the caller's pointer to it: call it as p^.delete(pSelf:=p).
	pSelf is cleared before the span is freed, so the caller never keeps a dangling pointer.
	A pointer to any other object is refused and left untouched, and nothing is released.
*)
METHOD delete : BOOL
VAR_IN_OUT
	pSelf: POINTER TO FB_Span;
END_VAR
VAR
	_pThis: POINTER TO FB_Span;
END_VAR
_pThis := THIS;
IF pSelf <> _pThis THEN
	RETURN;
END_IF

pSelf := 0;
__DELETE(_pThis);
delete := TRUE;
END_METHOD

//FB_Exit must be implemented explicitly. If there is an implementation, then the
//method is called before the controller removes the code of the function block instance
//(implicit call). The return value is not evaluated.
METHOD FB_Exit: BOOL
VAR_INPUT
    bInCopyCode: BOOL;  // TRUE: the exit method is called in order to leave the instance which will be copied afterwards (online change).
END_VAR
IF NOT bInCopyCode THEN
	THIS^.free();
END_IF
END_METHOD

(* Releases everything the span owns. Safe to call more than once. *)
METHOD free
IF THIS^.name <> 0 THEN THIS^.name^.delete(pSelf:=THIS^.name); END_IF
IF THIS^.traceId <> 0 THEN THIS^.traceId^.delete(pSelf:=THIS^.traceId); END_IF
IF THIS^.spanId <> 0 THEN THIS^.spanId^.delete(pSelf:=THIS^.spanId); END_IF
IF THIS^.traceState <> 0 THEN THIS^.traceState^.delete(pSelf:=THIS^.traceState); END_IF
IF THIS^.parentSpanId <> 0 THEN THIS^.parentSpanId^.delete(pSelf:=THIS^.parentSpanId); END_IF
IF THIS^.status <> 0 THEN THIS^.status^.delete(pSelf:=THIS^.status); END_IF
THIS^.attributes.free();
THIS^.links.free();
THIS^.scope.free();
THIS^.resource.free();
END_METHOD

(*
	Allocates a deep copy of this span, for a processor that keeps an ended span past onEnd.
	The copy owns copies of every member, so it stays valid after this span is released. This
	span is only read, apart from its links cursor. The caller owns pDest, which must be 0; on
	failure nothing is allocated and pDest is left alone.
*)
METHOD cloneTo : BOOL
VAR_IN_OUT
	pDest: POINTER TO FB_Span;
END_VAR
VAR_OUTPUT
	failureReason: E_SpanCloneFailureReason;
END_VAR
VAR
	_pClone: POINTER TO FB_Span;
	_pMessage: POINTER TO FB_String;
	_copied: BOOL;
	_attributesFailureReason: E_AttributesFailureReason;
	_linkFailureReason: E_LinkFailureReason;
END_VAR
cloneTo := FALSE;
failureReason := E_SpanCloneFailureReason.NA;

IF pDest <> 0 THEN
	failureReason := E_SpanCloneFailureReason.DESTINATION_ALREADY_ASSIGNED;
	RETURN;
END_IF

_pClone := __NEW(FB_Span);
IF _pClone = 0 THEN
	failureReason := E_SpanCloneFailureReason.MEMORY_ALLOCATION_FAILURE;
	RETURN;
END_IF

// the clone owns its members from here, so deleting it releases whatever was copied
_pClone^.kind := THIS^.kind;
_pClone^.startTimestamp := THIS^.startTimestamp;
_pClone^.endTimestamp := THIS^.endTimestamp;
_pClone^.flags := THIS^.flags;

_copied := (THIS^.name = 0 OR_ELSE ValueFactory.cloneString(
		pDest:=_pClone^.name,
		pSrc:=THIS^.name))
	AND_THEN (THIS^.traceId = 0 OR_ELSE ValueFactory.createTraceId(
		pDest:=_pClone^.traceId,
		pBytes:=ADR(THIS^.traceId^.bytes),
		nSize:=SIZEOF(THIS^.traceId^.bytes)))
	AND_THEN (THIS^.spanId = 0 OR_ELSE ValueFactory.createSpanId(
		pDest:=_pClone^.spanId,
		pBytes:=ADR(THIS^.spanId^.bytes),
		nSize:=SIZEOF(THIS^.spanId^.bytes)))
	AND_THEN (THIS^.parentSpanId = 0 OR_ELSE ValueFactory.createSpanId(
		pDest:=_pClone^.parentSpanId,
		pBytes:=ADR(THIS^.parentSpanId^.bytes),
		nSize:=SIZEOF(THIS^.parentSpanId^.bytes)))
	AND_THEN (THIS^.traceState = 0 OR_ELSE TraceStateFactory.clone(
		pDest:=_pClone^.traceState,
		pSrc:=THIS^.traceState))
	AND_THEN (THIS^.status = 0 OR_ELSE THIS^.status^.message = 0 OR_ELSE ValueFactory.cloneString(
		pDest:=_pMessage,
		pSrc:=THIS^.status^.message));
IF NOT _copied THEN
	IF _pMessage <> 0 THEN _pMessage^.delete(pSelf:=_pMessage); END_IF
	_pClone^.delete(pSelf:=_pClone);
	failureReason := E_SpanCloneFailureReason.VALUE_COPY_FAILURE;
	RETURN;
END_IF

IF THIS^.status <> 0 THEN
	_pClone^.status := __NEW(FB_Status(code:=THIS^.status^.code, message:=_pMessage));
	IF _pClone^.status = 0 THEN
		IF _pMessage <> 0 THEN _pMessage^.delete(pSelf:=_pMessage); END_IF
		_pClone^.delete(pSelf:=_pClone);
		failureReason := E_SpanCloneFailureReason.MEMORY_ALLOCATION_FAILURE;
		RETURN;
	END_IF
	_pMessage := 0;  // moved into the status
END_IF

IF NOT _pClone^.attributes.copyFrom(src:=THIS^.attributes, failureReason=>_attributesFailureReason) THEN
	_pClone^.delete(pSelf:=_pClone);
	IF _attributesFailureReason = E_AttributesFailureReason.MEMORY_ALLOCATION_FAILURE THEN
		failureReason := E_SpanCloneFailureReason.MEMORY_ALLOCATION_FAILURE;
	ELSE
		failureReason := E_SpanCloneFailureReason.ATTRIBUTE_COPY_FAILURE;
	END_IF
	RETURN;
END_IF

IF NOT _pClone^.links.copyFrom(src:=THIS^.links, failureReason=>_linkFailureReason) THEN
	_pClone^.delete(pSelf:=_pClone);
	IF _linkFailureReason = E_LinkFailureReason.MEMORY_ALLOCATION_FAILURE THEN
		failureReason := E_SpanCloneFailureReason.MEMORY_ALLOCATION_FAILURE;
	ELSE
		failureReason := E_SpanCloneFailureReason.LINK_COPY_FAILURE;
	END_IF
	RETURN;
END_IF

IF NOT _pClone^.resource.copyFrom(src:=THIS^.resource, failureResult=>_attributesFailureReason) THEN
	_pClone^.delete(pSelf:=_pClone);
	IF _attributesFailureReason = E_AttributesFailureReason.MEMORY_ALLOCATION_FAILURE THEN
		failureReason := E_SpanCloneFailureReason.MEMORY_ALLOCATION_FAILURE;
	ELSE
		failureReason := E_SpanCloneFailureReason.RESOURCE_COPY_FAILURE;
	END_IF
	RETURN;
END_IF

IF NOT _pClone^.scope.copyFrom(src:=THIS^.scope, failureResult=>_attributesFailureReason) THEN
	_pClone^.delete(pSelf:=_pClone);
	IF _attributesFailureReason = E_AttributesFailureReason.MEMORY_ALLOCATION_FAILURE THEN
		failureReason := E_SpanCloneFailureReason.MEMORY_ALLOCATION_FAILURE;
	ELSE
		failureReason := E_SpanCloneFailureReason.SCOPE_COPY_FAILURE;
	END_IF
	RETURN;
END_IF

// transfer ownership to the caller
pDest := _pClone;
_pClone := 0;
cloneTo := TRUE;
END_METHOD

(* TRUE when bit 0 of the trace flags, the W3C sampled flag, is set. *)
METHOD isSampled : BOOL
isSampled := (THIS^.flags AND 16#01) <> 0;
END_METHOD

(* Sets or clears bit 0 of the trace flags, the W3C sampled flag, and leaves the other bits. *)
METHOD setSampled
VAR_INPUT
	sampled: BOOL;
END_VAR
VAR CONSTANT
	TRACE_FLAG_SAMPLED: UDINT := 16#01;
END_VAR
IF sampled THEN
	THIS^.flags := THIS^.flags OR TRACE_FLAG_SAMPLED;
ELSE
	THIS^.flags := THIS^.flags AND NOT TRACE_FLAG_SAMPLED;
END_IF
END_METHOD

END_FUNCTION_BLOCK

// ---- OTEL/TRACING/TRACESTATE/FUNCTION_BLOCKS/FB_TraceState.TcPOU
(*
	Immutable W3C tracestate, created through TraceStateFactory and released with
	p^.delete(pSelf:=p). Holds the header in canonical form: its entries joined by ',', with
	optional whitespace and empty members removed. It always holds at least one valid entry,
	so no trace state is a 0 pointer, never an empty object. The string may be longer than
	T_MaxString: measure and copy it by length, never by assigning it to a STRING.
*)
{attribute 'enable_dynamic_creation'}
FUNCTION_BLOCK FB_TraceState
VAR
	_pString: POINTER TO STRING;
	_length: UDINT;
	_count: UDINT;
END_VAR

(*
	Releases this trace state and clears the caller's pointer to it: call it as p^.delete(pSelf:=p).
	pSelf is cleared before the trace state is freed, so the caller never keeps a dangling pointer.
	A pointer to any other object is refused and left untouched, and nothing is released.
*)
METHOD delete : BOOL
VAR_IN_OUT
	pSelf: POINTER TO FB_TraceState;
END_VAR
VAR
	_pThis: POINTER TO FB_TraceState;
END_VAR
_pThis := THIS;
IF pSelf <> _pThis THEN
	RETURN;
END_IF

pSelf := 0;
__DELETE(_pThis);
delete := TRUE;
END_METHOD

//FB_Exit must be implemented explicitly. If there is an implementation, then the
//method is called before the controller removes the code of the function block instance
//(implicit call). The return value is not evaluated.
METHOD FB_Exit: BOOL
VAR_INPUT
    bInCopyCode: BOOL;  // TRUE: the exit method is called in order to leave the instance which will be copied afterwards (online change).
END_VAR
// during an online change the copy keeps the string pointer, so it must not be released here
IF NOT bInCopyCode THEN
	THIS^.free();
END_IF
END_METHOD

//FB_Init is always available implicitly and it is used primarily for initialization.
//The return value is not evaluated. For a specific influence, you can also declare the
//methods explicitly and provide additional code there with the standard initialization
//code. You can evaluate the return value.
METHOD FB_Init: BOOL
VAR_INPUT
    bInitRetains: BOOL; // TRUE: the retain variables are initialized (reset warm / reset cold)
    bInCopyCode: BOOL;  // TRUE: the instance will be copied to the copy code afterward (online change)
	pString: POINTER TO STRING;  // canonical, null terminated; ownership transfers to the trace state
	length: UDINT;  // characters in pString, without the terminator
	count: UDINT;  // entries in pString
END_VAR
(*
Parsing, validation and allocation are done by TraceStateFactory and not the trace state
itself, that way a trace state is never allocated for a header that is not valid.
*)
THIS^._pString := pString;
THIS^._length := length;
THIS^._count := count;
FB_Init := TRUE;
END_METHOD

(*
	Releases the string. Safe to call more than once.
*)
METHOD free
IF THIS^._pString <> 0 THEN
	__DELETE(THIS^._pString);
	THIS^._pString := 0;
END_IF
THIS^._length := 0;
THIS^._count := 0;
END_METHOD

(* The number of entries. *)
PROPERTY count : UDINT
GET
count := THIS^._count;
END_GET
END_PROPERTY

(* The number of characters in the canonical string, without the terminator. *)
PROPERTY length : UDINT
GET
length := THIS^._length;
END_GET
END_PROPERTY

(* The canonical header string. Read only: the trace state owns it and never changes it. *)
PROPERTY pString : POINTER TO STRING
GET
pString := THIS^._pString;
END_GET
END_PROPERTY

END_FUNCTION_BLOCK

// ---- OTEL/TRACING/SPAN/FUNCTION_BLOCKS/FB_Status.TcPOU
{attribute 'enable_dynamic_creation'}
FUNCTION_BLOCK FB_Status
VAR_OUTPUT
	code: E_StatusCode;
	// optional and only set when status is an error. Owned by the status and released with it.
	message: POINTER TO FB_String;
END_VAR

(*
	Releases this status and clears the caller's pointer to it: call it as p^.delete(pSelf:=p).
	pSelf is cleared before the status is freed, so the caller never keeps a dangling pointer.
	A pointer to any other object is refused and left untouched, and nothing is released.
*)
METHOD delete : BOOL
VAR_IN_OUT
	pSelf: POINTER TO FB_Status;
END_VAR
VAR
	_pThis: POINTER TO FB_Status;
END_VAR
_pThis := THIS;
IF pSelf <> _pThis THEN
	RETURN;
END_IF

pSelf := 0;
__DELETE(_pThis);
delete := TRUE;
END_METHOD

//FB_Exit must be implemented explicitly. If there is an implementation, then the
//method is called before the controller removes the code of the function block instance
//(implicit call). The return value is not evaluated.
METHOD FB_Exit: BOOL
VAR_INPUT
    bInCopyCode: BOOL;  // TRUE: the exit method is called in order to leave the instance which will be copied afterwards (online change).  
END_VAR
THIS^.free();
END_METHOD

//FB_Init is always available implicitly and it is used primarily for initialization.
//The return value is not evaluated. For a specific influence, you can also declare the
//methods explicitly and provide additional code there with the standard initialization
//code. You can evaluate the return value.
METHOD FB_Init: BOOL
VAR_INPUT
    bInitRetains: BOOL; // TRUE: the retain variables are initialized (reset warm / reset cold)
    bInCopyCode: BOOL;  // TRUE: the instance will be copied to the copy code afterward (online change)
	code: E_StatusCode;
	message: POINTER TO FB_String;  // ownership transfers to the status; the creator clears its copy. 0 means none
END_VAR
THIS^.code := code;
THIS^.message := message;
END_METHOD

METHOD free
IF THIS^.message <> 0 THEN THIS^.message^.delete(pSelf:=THIS^.message); END_IF
END_METHOD

END_FUNCTION_BLOCK

// ---- OTEL/TRACING/LINK/FUNCTION_BLOCKS/FB_Links.TcPOU
(*
	The links of one span, oldest first. The collection owns every FB_Link it contains: push
	takes ownership and clears the caller's pointer, pop hands ownership back, and free
	releases what is left. The bound is maxCount, but never more than
	TcOtlp_GVL.MAX_LOOP_COUNT: a maxCount of zero, or one above that limit, is held to
	MAX_LOOP_COUNT so that free always reaches the end.
	reset and next walk the links without taking ownership, for readers such as serializers.
*)
FUNCTION_BLOCK FB_Links
VAR
	_head: POINTER TO ST_LinkedListNode;
	_tail: POINTER TO ST_LinkedListNode;
	_cursor: POINTER TO ST_LinkedListNode;  // next node returned by next; 0 at the end
END_VAR
VAR_OUTPUT
	count: UDINT;
	maxCount: UDINT;
	droppedCount: UDINT;  // links refused because the collection was full
END_VAR

(* The enforced bound: maxCount, held to MAX_LOOP_COUNT when it is zero or larger. *)
METHOD _capacity : UDINT
IF THIS^.maxCount = 0 OR THIS^.maxCount > TcOtlp_GVL.MAX_LOOP_COUNT THEN
	_capacity := TcOtlp_GVL.MAX_LOOP_COUNT;
ELSE
	_capacity := THIS^.maxCount;
END_IF
END_METHOD

METHOD FB_Exit : BOOL
VAR_INPUT
	bInCopyCode: BOOL;
END_VAR
IF NOT bInCopyCode THEN
	THIS^.free();
END_IF
END_METHOD

METHOD FB_Init : BOOL
VAR_INPUT
	bInitRetains: BOOL;
	bInCopyCode: BOOL;
	maxCount: UDINT := TcOtlp_GVL.DEFAULT_MAX_LINK_COUNT;
END_VAR
THIS^.maxCount := maxCount;
END_METHOD

(*
	Releases every owned link and clears droppedCount. push holds count to MAX_LOOP_COUNT, so
	the loop always reaches the end. If it ever stops early, the unreleased nodes stay in the
	collection and free returns FALSE, so a later call can finish the job.
*)
METHOD free : BOOL
VAR
	_idx: UDINT;
	_node: POINTER TO ST_LinkedListNode;
	_link: POINTER TO FB_Link;
END_VAR
FOR _idx := 0 TO TcOtlp_GVL.MAX_LOOP_COUNT DO
	IF THIS^._head = 0 THEN
		EXIT;
	END_IF

	_node := THIS^._head;
	THIS^._head := _node^.nxt;
	IF _node^.val <> 0 THEN
		_link := _node^.val;
		_node^.val := 0;
		_link^.delete(pSelf:=_link);
	END_IF
	__DELETE(_node);
	_node := 0;
	IF THIS^.count > 0 THEN
		THIS^.count := THIS^.count - 1;
	END_IF
END_FOR

IF THIS^._head = 0 THEN
	THIS^._tail := 0;
	THIS^.count := 0;
	THIS^.droppedCount := 0;
END_IF
THIS^._cursor := THIS^._head;
free := THIS^._head = 0;
END_METHOD

(*
	Returns the link at the cursor and advances it, or 0 after the last link. The link is
	borrowed: the collection still owns it, and it is valid only until it is popped or freed.
	Call reset first.
*)
METHOD next : POINTER TO FB_Link
next := 0;
IF THIS^._cursor <> 0 THEN
	next := THIS^._cursor^.val;
	THIS^._cursor := THIS^._cursor^.nxt;
END_IF
END_METHOD

(* Moves the oldest link to pValue, which must be 0. The caller owns it on success. *)
METHOD pop : BOOL
VAR_IN_OUT
	pValue: POINTER TO FB_Link;
END_VAR
VAR_OUTPUT
	failureReason: E_LinkFailureReason;
END_VAR
VAR
	_node: POINTER TO ST_LinkedListNode;
END_VAR
pop := FALSE;
failureReason := E_LinkFailureReason.NA;

IF pValue <> 0 THEN
	failureReason := E_LinkFailureReason.DESTINATION_ALREADY_ASSIGNED;
	RETURN;
END_IF
IF THIS^._head = 0 THEN
	failureReason := E_LinkFailureReason.LINKS_EMPTY;
	RETURN;
END_IF

_node := THIS^._head;
THIS^._head := _node^.nxt;
IF THIS^._head = 0 THEN
	THIS^._tail := 0;
END_IF
IF THIS^._cursor = _node THEN
	THIS^._cursor := THIS^._head;
END_IF

pValue := _node^.val;
_node^.val := 0;
_node^.nxt := 0;
__DELETE(_node);
_node := 0;
THIS^.count := THIS^.count - 1;
pop := failureReason = E_LinkFailureReason.NA;
END_METHOD

(*
	Takes ownership of the link and clears pValue. On failure pValue is left unchanged and
	still owned by the caller. A full collection keeps the links it has, as the OpenTelemetry
	limits require: the new link is refused with LINK_COUNT_LIMIT_REACHED and counted in
	droppedCount, and the caller releases it.
*)
METHOD push : BOOL
VAR_IN_OUT
	pValue: POINTER TO FB_Link;
END_VAR
VAR_OUTPUT
	failureReason: E_LinkFailureReason;
END_VAR
VAR
	_node: POINTER TO ST_LinkedListNode;
END_VAR
push := FALSE;
failureReason := E_LinkFailureReason.NA;

IF pValue = 0 THEN
	failureReason := E_LinkFailureReason.LINK_POINTER_NULL;
	RETURN;
END_IF

IF THIS^.count >= THIS^._capacity() THEN
	failureReason := E_LinkFailureReason.LINK_COUNT_LIMIT_REACHED;
	THIS^.droppedCount := THIS^.droppedCount + 1;
	RETURN;
END_IF

_node := __NEW(ST_LinkedListNode);
IF _node = 0 THEN
	failureReason := E_LinkFailureReason.MEMORY_ALLOCATION_FAILURE;
	RETURN;
END_IF

_node^.val := pValue;
_node^.nxt := 0;
IF THIS^._tail = 0 THEN
	THIS^._head := _node;
	THIS^._cursor := _node;
ELSE
	THIS^._tail^.nxt := _node;
END_IF
THIS^._tail := _node;
THIS^.count := THIS^.count + 1;
pValue := 0;
push := failureReason = E_LinkFailureReason.NA;
END_METHOD

(* Moves the cursor to the oldest link, so next starts from the head. *)
METHOD reset
THIS^._cursor := THIS^._head;
END_METHOD

(*
	Adds a copy of every link in src, oldest first, through LinkFactory.fromLink, and carries
	src's droppedCount over. src is only read, apart from its cursor. On failure the links
	copied so far stay in this collection, for the caller to release.
*)
METHOD copyFrom : BOOL
VAR_IN_OUT
	src: FB_Links;
END_VAR
VAR_OUTPUT
	failureReason: E_LinkFailureReason;
END_VAR
VAR
	_idx: UDINT;
	_pLink: POINTER TO FB_Link;
END_VAR
copyFrom := FALSE;
failureReason := E_LinkFailureReason.NA;

THIS^.droppedCount := THIS^.droppedCount + src.droppedCount;

// src.count never exceeds MAX_LOOP_COUNT, so this loop is bounded
src.reset();
FOR _idx := 1 TO src.count DO
	IF NOT LinkFactory.fromLink(pDest:=_pLink, pSrc:=src.next(), failureReason=>failureReason)
		OR_ELSE NOT THIS^.push(pValue:=_pLink, failureReason=>failureReason) THEN
		IF _pLink <> 0 THEN _pLink^.delete(pSelf:=_pLink); END_IF
		RETURN;
	END_IF
END_FOR

copyFrom := TRUE;
END_METHOD

END_FUNCTION_BLOCK

// ---- OTEL/TRACING/LINK/FUNCTION_BLOCKS/FB_Link.TcPOU
(*
	A pointer from one span to another span's context, possibly in another trace. Build it
	through LinkFactory, which validates the context and copies its identity.
	The link owns every pointer member and releases them in free.
*)
{attribute 'enable_dynamic_creation'}
FUNCTION_BLOCK FB_Link
VAR_INPUT
	// written by LinkFactory
	traceId: POINTER TO FB_TraceId;
	spanId: POINTER TO FB_SpanId;
	traceState: POINTER TO FB_TraceState;  // optional; 0 means none

	// the linked context's trace flags and remoteness; see E_SpanFlags
	flags: UDINT;
END_VAR
VAR_OUTPUT
	attributes: FB_Attributes(maxCount := TcOtlp_GVL.DEFAULT_MAX_ATTRIBUTE_COUNT);
END_VAR

(*
	Releases this link and clears the caller's pointer to it: call it as p^.delete(pSelf:=p).
	pSelf is cleared before the link is freed, so the caller never keeps a dangling pointer.
	A pointer to any other object is refused and left untouched, and nothing is released.
*)
METHOD delete : BOOL
VAR_IN_OUT
	pSelf: POINTER TO FB_Link;
END_VAR
VAR
	_pThis: POINTER TO FB_Link;
END_VAR
_pThis := THIS;
IF pSelf <> _pThis THEN
	RETURN;
END_IF

pSelf := 0;
__DELETE(_pThis);
delete := TRUE;
END_METHOD

//FB_Exit must be implemented explicitly. If there is an implementation, then the
//method is called before the controller removes the code of the function block instance
//(implicit call). The return value is not evaluated.
METHOD FB_Exit: BOOL
VAR_INPUT
    bInCopyCode: BOOL;  // TRUE: the exit method is called in order to leave the instance which will be copied afterwards (online change).  
END_VAR
IF NOT bInCopyCode THEN
	THIS^.free();
END_IF
END_METHOD

//FB_Init is always available implicitly and it is used primarily for initialization.
//The return value is not evaluated. For a specific influence, you can also declare the
//methods explicitly and provide additional code there with the standard initialization
//code. You can evaluate the return value.
METHOD FB_Init: BOOL
VAR_INPUT
    bInitRetains: BOOL; // TRUE: the retain variables are initialized (reset warm / reset cold)
    bInCopyCode: BOOL;  // TRUE: the instance will be copied to the copy code afterward (online change)   
END_VAR
END_METHOD

(*
	Releases every value the link owns and clears the pointers. Safe to call more than once.
*)
METHOD free
IF THIS^.traceId <> 0 THEN THIS^.traceId^.delete(pSelf:=THIS^.traceId); END_IF
IF THIS^.spanId <> 0 THEN THIS^.spanId^.delete(pSelf:=THIS^.spanId); END_IF
IF THIS^.traceState <> 0 THEN THIS^.traceState^.delete(pSelf:=THIS^.traceState); END_IF
THIS^.attributes.free();
THIS^.flags := 0;
END_METHOD

END_FUNCTION_BLOCK

// ---- OTEL/TRACING/LINK/FUNCTION_BLOCKS/LinkFactory.TcPOU
(*
	Creates FB_Link values and keeps their invariants: a link always points at a valid span
	context and owns copies of its identity. Attributes can be added to the link's attributes
	after it is created.
*)
PROGRAM LinkFactory

(*
	Allocates a link to the given span context. The context is borrowed: the link holds copies
	of its trace id, span id and trace state, so it stays valid after the context is released.
	The link's flags carry the context's trace flags and remoteness. The caller owns pDest,
	which must be 0; on failure nothing is allocated and pDest is left alone.
*)
METHOD fromContext : BOOL
VAR_IN_OUT
	pDest: POINTER TO FB_Link;
END_VAR
VAR_INPUT
	pContext: POINTER TO FB_SpanContext;
END_VAR
VAR_OUTPUT
	failureReason: E_LinkFailureReason;
END_VAR
VAR
	_ctxTraceId: REFERENCE TO FB_TraceId;
	_ctxSpanId: REFERENCE TO FB_SpanId;
	_pNew: POINTER TO FB_Link;
	_copied: BOOL;
	_flags: UDINT;
END_VAR
fromContext := FALSE;
failureReason := E_LinkFailureReason.NA;

IF pDest <> 0 THEN
	failureReason := E_LinkFailureReason.DESTINATION_ALREADY_ASSIGNED;
	RETURN;
END_IF
IF pContext = 0 THEN
	failureReason := E_LinkFailureReason.CONTEXT_POINTER_NULL;
	RETURN;
END_IF
IF NOT pContext^.isValid() THEN
	failureReason := E_LinkFailureReason.CONTEXT_INVALID;
	RETURN;
END_IF

_pNew := __NEW(FB_Link);
IF _pNew = 0 THEN
	failureReason := E_LinkFailureReason.MEMORY_ALLOCATION_FAILURE;
	RETURN;
END_IF

// the link owns its members from here, so deleting it releases whatever was copied
_ctxTraceId REF= pContext^.traceId;
_ctxSpanId REF= pContext^.spanId;
_copied := ValueFactory.createTraceId(
		pDest:=_pNew^.traceId,
		pBytes:=ADR(_ctxTraceId.bytes),
		nSize:=SIZEOF(_ctxTraceId.bytes))
	AND_THEN ValueFactory.createSpanId(
		pDest:=_pNew^.spanId,
		pBytes:=ADR(_ctxSpanId.bytes),
		nSize:=SIZEOF(_ctxSpanId.bytes))
	AND_THEN (pContext^.traceState = 0 OR_ELSE TraceStateFactory.clone(
		pDest:=_pNew^.traceState,
		pSrc:=pContext^.traceState));
IF NOT _copied THEN
	_pNew^.delete(pSelf:=_pNew);
	failureReason := E_LinkFailureReason.MEMORY_ALLOCATION_FAILURE;
	RETURN;
END_IF

// the same encoding a span uses for its parent: trace flags plus known remoteness
_flags := (pContext^.traceFlags AND TO_UDINT(E_SpanFlags.SPAN_FLAGS_TRACE_FLAGS_MASK))
	OR TO_UDINT(E_SpanFlags.SPAN_FLAGS_CONTEXT_HAS_IS_REMOTE_MASK);
IF pContext^.isRemote() THEN
	_flags := _flags OR TO_UDINT(E_SpanFlags.SPAN_FLAGS_CONTEXT_IS_REMOTE_MASK);
END_IF
_pNew^.flags := _flags;

// transfer ownership to the caller
pDest := _pNew;
_pNew := 0;
fromContext := TRUE;
END_METHOD

(*
	Allocates a link to a span the caller holds, such as a running or ended span in this PLC.
	The span is borrowed and unchanged. The link is built from the span's context, so it is
	local: remoteness is known and not remote. The caller owns pDest, which must be 0.
*)
METHOD fromSpan : BOOL
VAR_IN_OUT
	pDest: POINTER TO FB_Link;
END_VAR
VAR_INPUT
	pSpan: POINTER TO FB_Span;
END_VAR
VAR_OUTPUT
	failureReason: E_LinkFailureReason;
END_VAR
VAR
	_pContext: POINTER TO FB_SpanContext;
END_VAR
fromSpan := FALSE;
failureReason := E_LinkFailureReason.NA;

IF pDest <> 0 THEN
	failureReason := E_LinkFailureReason.DESTINATION_ALREADY_ASSIGNED;
	RETURN;
END_IF
IF pSpan = 0 THEN
	failureReason := E_LinkFailureReason.SPAN_POINTER_NULL;
	RETURN;
END_IF
IF pSpan^.traceId = 0 OR pSpan^.spanId = 0 THEN
	failureReason := E_LinkFailureReason.CONTEXT_INVALID;
	RETURN;
END_IF

IF NOT ContextFactory.fromSpan(pDest:=_pContext, pSpan:=pSpan) THEN
	IF _pContext <> 0 THEN _pContext^.delete(pSelf:=_pContext); END_IF
	failureReason := E_LinkFailureReason.MEMORY_ALLOCATION_FAILURE;
	RETURN;
END_IF
fromSpan := LinkFactory.fromContext(pDest:=pDest, pContext:=_pContext, failureReason=>failureReason);
_pContext^.delete(pSelf:=_pContext);
END_METHOD

(*
	Allocates a copy of a link, for a span copy that must outlive the original. The source is
	borrowed and unchanged. The copy owns its own identity, trace state and attributes. The
	caller owns pDest, which must be 0; on failure nothing is allocated and pDest is left alone.
*)
METHOD fromLink : BOOL
VAR_IN_OUT
	pDest: POINTER TO FB_Link;
END_VAR
VAR_INPUT
	pSrc: POINTER TO FB_Link;
END_VAR
VAR_OUTPUT
	failureReason: E_LinkFailureReason;
END_VAR
VAR
	_pNew: POINTER TO FB_Link;
	_copied: BOOL;
	_attributesFailureReason: E_AttributesFailureReason;
END_VAR
fromLink := FALSE;
failureReason := E_LinkFailureReason.NA;

IF pDest <> 0 THEN
	failureReason := E_LinkFailureReason.DESTINATION_ALREADY_ASSIGNED;
	RETURN;
END_IF
IF pSrc = 0 THEN
	failureReason := E_LinkFailureReason.LINK_POINTER_NULL;
	RETURN;
END_IF
IF pSrc^.traceId = 0 OR pSrc^.spanId = 0 THEN
	failureReason := E_LinkFailureReason.CONTEXT_INVALID;
	RETURN;
END_IF

_pNew := __NEW(FB_Link);
IF _pNew = 0 THEN
	failureReason := E_LinkFailureReason.MEMORY_ALLOCATION_FAILURE;
	RETURN;
END_IF

// the copy owns its members from here, so deleting it releases whatever was copied
_copied := ValueFactory.createTraceId(
		pDest:=_pNew^.traceId,
		pBytes:=ADR(pSrc^.traceId^.bytes),
		nSize:=SIZEOF(pSrc^.traceId^.bytes))
	AND_THEN ValueFactory.createSpanId(
		pDest:=_pNew^.spanId,
		pBytes:=ADR(pSrc^.spanId^.bytes),
		nSize:=SIZEOF(pSrc^.spanId^.bytes))
	AND_THEN (pSrc^.traceState = 0 OR_ELSE TraceStateFactory.clone(
		pDest:=_pNew^.traceState,
		pSrc:=pSrc^.traceState));
IF NOT _copied THEN
	_pNew^.delete(pSelf:=_pNew);
	failureReason := E_LinkFailureReason.MEMORY_ALLOCATION_FAILURE;
	RETURN;
END_IF
_pNew^.flags := pSrc^.flags;

IF NOT _pNew^.attributes.copyFrom(src:=pSrc^.attributes, failureReason=>_attributesFailureReason) THEN
	_pNew^.delete(pSelf:=_pNew);
	IF _attributesFailureReason = E_AttributesFailureReason.MEMORY_ALLOCATION_FAILURE THEN
		failureReason := E_LinkFailureReason.MEMORY_ALLOCATION_FAILURE;
	ELSE
		failureReason := E_LinkFailureReason.ATTRIBUTE_COPY_FAILURE;
	END_IF
	RETURN;
END_IF

// transfer ownership to the caller
pDest := _pNew;
_pNew := 0;
fromLink := TRUE;
END_METHOD

END_PROGRAM

// ---- OTEL/TRACING/SPAN/FUNCTION_BLOCKS/FB_SpanContext.TcPOU
(*
	Immutable snapshot of the identity of one span, created through ContextFactory.buildContext.
	The identifiers are copies, so a context stays valid after the span it came from has ended.
*)
{attribute 'enable_dynamic_creation'}
FUNCTION_BLOCK FB_SpanContext
VAR
	_traceId: FB_TraceId;
	_spanId: FB_SpanId;
	_traceState: POINTER TO FB_TraceState;
	_traceFlags: UDINT;
END_VAR

METHOD _isZero : BOOL
VAR_INPUT
	pBytes: POINTER TO BYTE;
	size: UDINT;
END_VAR
VAR
	i: UDINT;
END_VAR
// bounded by the width of an identifier, at most 16 bytes
_isZero := TRUE;
WHILE i < size DO
	IF pBytes[i] <> 0 THEN
		_isZero := FALSE;
		RETURN;
	END_IF
	i := i + 1;
END_WHILE
END_METHOD

(*
	Releases this context and clears the caller's pointer to it: call it as p^.delete(pSelf:=p).
	pSelf is cleared before the context is freed, so the caller never keeps a dangling pointer.
	A pointer to any other object is refused and left untouched, and nothing is released.
*)
METHOD delete : BOOL
VAR_IN_OUT
	pSelf: POINTER TO FB_SpanContext;
END_VAR
VAR
	_pThis: POINTER TO FB_SpanContext;
END_VAR
_pThis := THIS;
IF pSelf <> _pThis THEN
	RETURN;
END_IF

pSelf := 0;
__DELETE(_pThis);
delete := TRUE;
END_METHOD

//FB_Exit must be implemented explicitly. If there is an implementation, then the
//method is called before the controller removes the code of the function block instance
//(implicit call). The return value is not evaluated.
METHOD FB_Exit: BOOL
VAR_INPUT
    bInCopyCode: BOOL;  // TRUE: the exit method is called in order to leave the instance which will be copied afterwards (online change).
END_VAR
// during an online change the copy keeps the trace state pointer, so it must not be released here
IF NOT bInCopyCode THEN
	THIS^.free();
END_IF
END_METHOD

//FB_Init is always available implicitly and it is used primarily for initialization.
//The return value is not evaluated. For a specific influence, you can also declare the
//methods explicitly and provide additional code there with the standard initialization
//code. You can evaluate the return value.
METHOD FB_Init: BOOL
VAR_INPUT
    bInitRetains: BOOL; // TRUE: the retain variables are initialized (reset warm / reset cold)
    bInCopyCode: BOOL;  // TRUE: the instance will be copied to the copy code afterward (online change)
	pTraceId: POINTER TO FB_TraceId;  // copied
	pSpanId: POINTER TO FB_SpanId;  // copied
	pTraceState: POINTER TO FB_TraceState;  // ownership transfers to the context; 0 means none
	traceFlags: UDINT;
END_VAR
(*
Allocation and argument checks are done by ContextFactory and not the context itself,
that way a new context never gets allocated if building it fails.
The identity is not validated; producers are responsible for what they build.
*)
IF pTraceId <> 0 THEN
	MEMCPY(ADR(THIS^._traceId.bytes), ADR(pTraceId^.bytes), SIZEOF(THIS^._traceId.bytes));
END_IF
IF pSpanId <> 0 THEN
	MEMCPY(ADR(THIS^._spanId.bytes), ADR(pSpanId^.bytes), SIZEOF(THIS^._spanId.bytes));
END_IF
THIS^._traceState := pTraceState;
THIS^._traceFlags := traceFlags;
FB_Init := TRUE;
END_METHOD

//FB_Reinit is called after the instance has been copied during an online change.
//The return value is not evaluated.
METHOD FB_Reinit: BOOL
// nothing to fix up: the trace state lives on the heap and does not move with the instance,
// and no member points back into this instance
FB_Reinit := TRUE;
END_METHOD

(*
	Releases the trace state and clears the identity. Safe to call more than once.
*)
METHOD free
IF THIS^._traceState <> 0 THEN
	THIS^._traceState^.delete(pSelf:=THIS^._traceState);
END_IF
THIS^._traceId.free();
THIS^._spanId.free();
THIS^._traceFlags := 0;
END_METHOD

(*
	TRUE only when remoteness is known and the span is remote, meaning the context was
	extracted from a carrier rather than produced by a local tracer.
	FALSE covers both "known local" and "not known".
*)
METHOD isRemote : BOOL
isRemote := (THIS^._traceFlags AND TO_UDINT(E_SpanFlags.SPAN_FLAGS_CONTEXT_HAS_IS_REMOTE_MASK)) <> 0
	AND (THIS^._traceFlags AND TO_UDINT(E_SpanFlags.SPAN_FLAGS_CONTEXT_IS_REMOTE_MASK)) <> 0;
END_METHOD

(*
	TRUE if and only if both the trace ID and the span ID are non-zero.
*)
METHOD isValid : BOOL
isValid := NOT THIS^._isZero(pBytes := ADR(THIS^._traceId.bytes), size := SIZEOF(THIS^._traceId.bytes))
	AND NOT THIS^._isZero(pBytes := ADR(THIS^._spanId.bytes), size := SIZEOF(THIS^._spanId.bytes));
END_METHOD

PROPERTY spanId : REFERENCE TO FB_SpanId
GET
spanId REF= THIS^._spanId;
END_GET
END_PROPERTY

PROPERTY traceFlags : UDINT
GET
traceFlags := THIS^._traceFlags;
END_GET
END_PROPERTY

PROPERTY traceId : REFERENCE TO FB_TraceId
GET
traceId REF= THIS^._traceId;
END_GET
END_PROPERTY

// borrowed; 0 when the context carries no trace state. The context owns and releases it.
PROPERTY traceState : POINTER TO FB_TraceState
GET
traceState := THIS^._traceState;
END_GET
END_PROPERTY

END_FUNCTION_BLOCK

